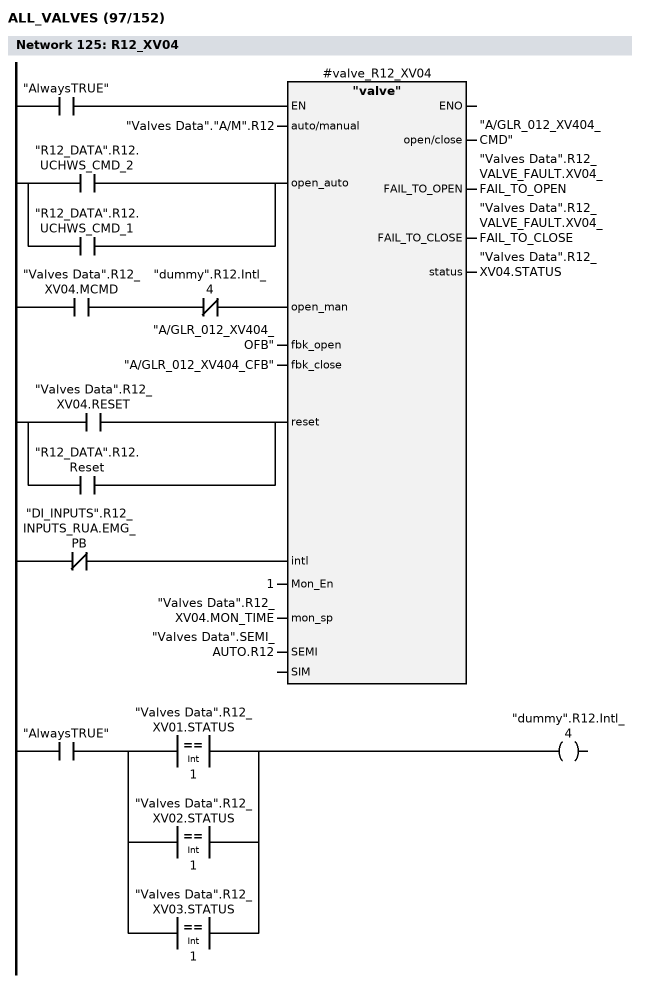
   RUNG wire#powerrail
      Contact( "AlwaysTRUE" )
      #valve_R12_XV04(open_auto := wire#w1, open_man := wire#w2, reset := wire#w3, intl := wire#w4, "auto/manual" := "Valves Data"."A/M".R12, fbk_open := "A/GLR_012_XV404_OFB", fbk_close := "A/GLR_012_XV404_CFB", Mon_En := 1, mon_sp := "Valves Data".R12_XV04.MON_TIME, SEMI := "Valves Data".SEMI_AUTO.R12, SIM :=, "open/close" => "A/GLR_012_XV404_CMD", FAIL_TO_OPEN => "Valves Data".R12_VALVE_FAULT.XV04_FAIL_TO_OPEN, FAIL_TO_CLOSE => "Valves Data".R12_VALVE_FAULT.XV04_FAIL_TO_CLOSE, status => "Valves Data".R12_XV04.STATUS)
   END_RUNG
   RUNG wire#powerrail
      Contact( "R12_DATA".R12.UCHWS_CMD_2 )
   END_RUNG wire#w1
   RUNG wire#powerrail
      Contact( "R12_DATA".R12.UCHWS_CMD_1 )
   END_RUNG wire#w1
   RUNG wire#powerrail
      Contact( "Valves Data".R12_XV04.MCMD )
      I_Contact( "dummy".R12.Intl_4 )
   END_RUNG wire#w2
   RUNG wire#powerrail
      Contact( "Valves Data".R12_XV04.RESET )
   END_RUNG wire#w3
   RUNG wire#powerrail
      Contact( "R12_DATA".R12.Reset )
   END_RUNG wire#w3
   RUNG wire#powerrail
      I_Contact( "DI_INPUTS".R12_INPUTS_RUA.EMG_PB )
   END_RUNG wire#w4
   RUNG wire#powerrail
      Contact( "AlwaysTRUE" )
      wire#w5
      { S7_Templates := "SrcType := Int" } EQ_Contact(in1 := "Valves Data".R12_XV01.STATUS, in2 := 1)
      wire#w6
      Coil( "dummy".R12.Intl_4 )
   END_RUNG
   RUNG wire#w5
      { S7_Templates := "SrcType := Int" } EQ_Contact(in1 := "Valves Data".R12_XV02.STATUS, in2 := 1)
   END_RUNG wire#w6
   RUNG wire#w5
      { S7_Templates := "SrcType := Int" } EQ_Contact(in1 := "Valves Data".R12_XV03.STATUS, in2 := 1)
   END_RUNG wire#w6
   // the same network as SCL:
   IF "AlwaysTRUE" THEN
       #valve_R12_XV04("auto/manual" := "Valves Data"."A/M".R12,   // "valve"
                       open_auto := "R12_DATA".R12.UCHWS_CMD_2 OR "R12_DATA".R12.UCHWS_CMD_1,
                       open_man := "Valves Data".R12_XV04.MCMD AND NOT "dummy".R12.Intl_4,
                       fbk_open := "A/GLR_012_XV404_OFB",
                       fbk_close := "A/GLR_012_XV404_CFB",
                       reset := "Valves Data".R12_XV04.RESET OR "R12_DATA".R12.Reset,
                       intl := NOT "DI_INPUTS".R12_INPUTS_RUA.EMG_PB,
                       Mon_En := 1,
                       mon_sp := "Valves Data".R12_XV04.MON_TIME,
                       SEMI := "Valves Data".SEMI_AUTO.R12,
                       "open/close" => "A/GLR_012_XV404_CMD",
                       FAIL_TO_OPEN => "Valves Data".R12_VALVE_FAULT.XV04_FAIL_TO_OPEN,
                       FAIL_TO_CLOSE => "Valves Data".R12_VALVE_FAULT.XV04_FAIL_TO_CLOSE,
                       status => "Valves Data".R12_XV04.STATUS);
   END_IF;
   "dummy".R12.Intl_4 := "AlwaysTRUE" AND (("Valves Data".R12_XV01.STATUS = 1) OR ("Valves Data".R12_XV02.STATUS = 1) OR ("Valves Data".R12_XV03.STATUS = 1));
END_REGION

REGION Network 126: R12_XV05
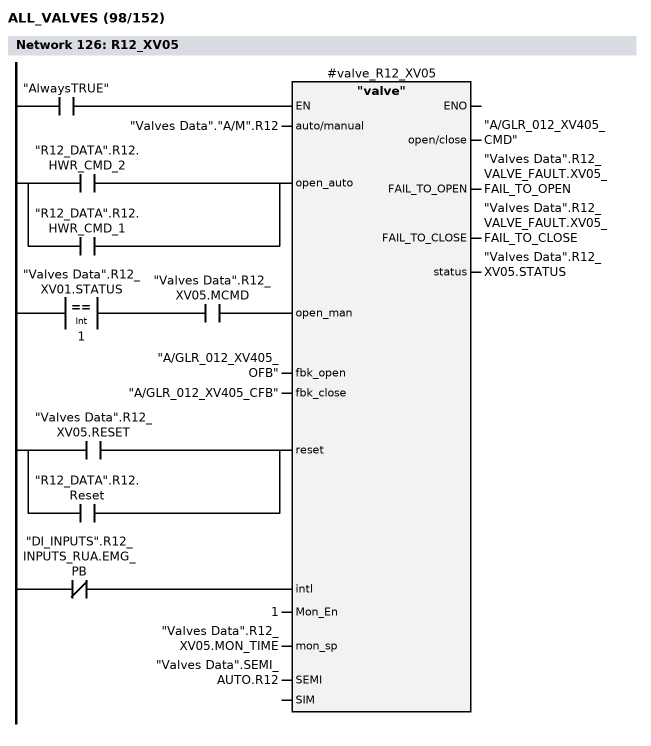
   RUNG wire#powerrail
      Contact( "AlwaysTRUE" )
      #valve_R12_XV05(open_auto := wire#w1, open_man := wire#w2, reset := wire#w3, intl := wire#w4, "auto/manual" := "Valves Data"."A/M".R12, fbk_open := "A/GLR_012_XV405_OFB", fbk_close := "A/GLR_012_XV405_CFB", Mon_En := 1, mon_sp := "Valves Data".R12_XV05.MON_TIME, SEMI := "Valves Data".SEMI_AUTO.R12, SIM :=, "open/close" => "A/GLR_012_XV405_CMD", FAIL_TO_OPEN => "Valves Data".R12_VALVE_FAULT.XV05_FAIL_TO_OPEN, FAIL_TO_CLOSE => "Valves Data".R12_VALVE_FAULT.XV05_FAIL_TO_CLOSE, status => "Valves Data".R12_XV05.STATUS)
   END_RUNG
   RUNG wire#powerrail
      Contact( "R12_DATA".R12.HWR_CMD_2 )
   END_RUNG wire#w1
   RUNG wire#powerrail
      Contact( "R12_DATA".R12.HWR_CMD_1 )
   END_RUNG wire#w1
   RUNG wire#powerrail
      { S7_Templates := "SrcType := Int" } EQ_Contact(in1 := "Valves Data".R12_XV01.STATUS, in2 := 1)
      Contact( "Valves Data".R12_XV05.MCMD )
   END_RUNG wire#w2
   RUNG wire#powerrail
      Contact( "Valves Data".R12_XV05.RESET )
   END_RUNG wire#w3
   RUNG wire#powerrail
      Contact( "R12_DATA".R12.Reset )
   END_RUNG wire#w3
   RUNG wire#powerrail
      I_Contact( "DI_INPUTS".R12_INPUTS_RUA.EMG_PB )
   END_RUNG wire#w4
   // the same network as SCL:
   IF "AlwaysTRUE" THEN
       #valve_R12_XV05("auto/manual" := "Valves Data"."A/M".R12,   // "valve"
                       open_auto := "R12_DATA".R12.HWR_CMD_2 OR "R12_DATA".R12.HWR_CMD_1,
                       open_man := ("Valves Data".R12_XV01.STATUS = 1) AND "Valves Data".R12_XV05.MCMD,
                       fbk_open := "A/GLR_012_XV405_OFB",
                       fbk_close := "A/GLR_012_XV405_CFB",
                       reset := "Valves Data".R12_XV05.RESET OR "R12_DATA".R12.Reset,
                       intl := NOT "DI_INPUTS".R12_INPUTS_RUA.EMG_PB,
                       Mon_En := 1,
                       mon_sp := "Valves Data".R12_XV05.MON_TIME,
                       SEMI := "Valves Data".SEMI_AUTO.R12,
                       "open/close" => "A/GLR_012_XV405_CMD",
                       FAIL_TO_OPEN => "Valves Data".R12_VALVE_FAULT.XV05_FAIL_TO_OPEN,
                       FAIL_TO_CLOSE => "Valves Data".R12_VALVE_FAULT.XV05_FAIL_TO_CLOSE,
                       status => "Valves Data".R12_XV05.STATUS);
   END_IF;
END_REGION

REGION Network 127: R12_XV06
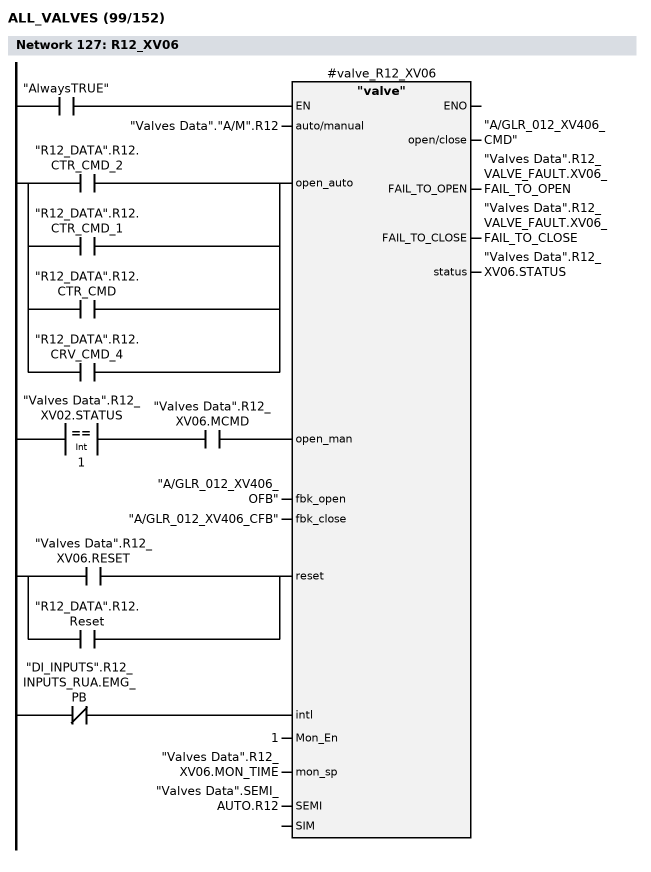
   RUNG wire#powerrail
      Contact( "AlwaysTRUE" )
      #valve_R12_XV06(open_auto := wire#w1, open_man := wire#w2, reset := wire#w3, intl := wire#w4, "auto/manual" := "Valves Data"."A/M".R12, fbk_open := "A/GLR_012_XV406_OFB", fbk_close := "A/GLR_012_XV406_CFB", Mon_En := 1, mon_sp := "Valves Data".R12_XV06.MON_TIME, SEMI := "Valves Data".SEMI_AUTO.R12, SIM :=, "open/close" => "A/GLR_012_XV406_CMD", FAIL_TO_OPEN => "Valves Data".R12_VALVE_FAULT.XV06_FAIL_TO_OPEN, FAIL_TO_CLOSE => "Valves Data".R12_VALVE_FAULT.XV06_FAIL_TO_CLOSE, status => "Valves Data".R12_XV06.STATUS)
   END_RUNG
   RUNG wire#powerrail
      Contact( "R12_DATA".R12.CTR_CMD_2 )
   END_RUNG wire#w1
   RUNG wire#powerrail
      Contact( "R12_DATA".R12.CTR_CMD_1 )
   END_RUNG wire#w1
   RUNG wire#powerrail
      Contact( "R12_DATA".R12.CTR_CMD )
   END_RUNG wire#w1
   RUNG wire#powerrail
      Contact( "R12_DATA".R12.CRV_CMD_4 )
   END_RUNG wire#w1
   RUNG wire#powerrail
      { S7_Templates := "SrcType := Int" } EQ_Contact(in1 := "Valves Data".R12_XV02.STATUS, in2 := 1)
      Contact( "Valves Data".R12_XV06.MCMD )
   END_RUNG wire#w2
   RUNG wire#powerrail
      Contact( "Valves Data".R12_XV06.RESET )
   END_RUNG wire#w3
   RUNG wire#powerrail
      Contact( "R12_DATA".R12.Reset )
   END_RUNG wire#w3
   RUNG wire#powerrail
      I_Contact( "DI_INPUTS".R12_INPUTS_RUA.EMG_PB )
   END_RUNG wire#w4
   // the same network as SCL:
   IF "AlwaysTRUE" THEN
       #valve_R12_XV06("auto/manual" := "Valves Data"."A/M".R12,   // "valve"
                       open_auto := "R12_DATA".R12.CTR_CMD_2 OR "R12_DATA".R12.CTR_CMD_1 OR "R12_DATA".R12.CTR_CMD OR "R12_DATA".R12.CRV_CMD_4,
                       open_man := ("Valves Data".R12_XV02.STATUS = 1) AND "Valves Data".R12_XV06.MCMD,
                       fbk_open := "A/GLR_012_XV406_OFB",
                       fbk_close := "A/GLR_012_XV406_CFB",
                       reset := "Valves Data".R12_XV06.RESET OR "R12_DATA".R12.Reset,
                       intl := NOT "DI_INPUTS".R12_INPUTS_RUA.EMG_PB,
                       Mon_En := 1,
                       mon_sp := "Valves Data".R12_XV06.MON_TIME,
                       SEMI := "Valves Data".SEMI_AUTO.R12,
                       "open/close" => "A/GLR_012_XV406_CMD",
                       FAIL_TO_OPEN => "Valves Data".R12_VALVE_FAULT.XV06_FAIL_TO_OPEN,
                       FAIL_TO_CLOSE => "Valves Data".R12_VALVE_FAULT.XV06_FAIL_TO_CLOSE,
                       status => "Valves Data".R12_XV06.STATUS);
   END_IF;
END_REGION

REGION Network 128: R12_XV07
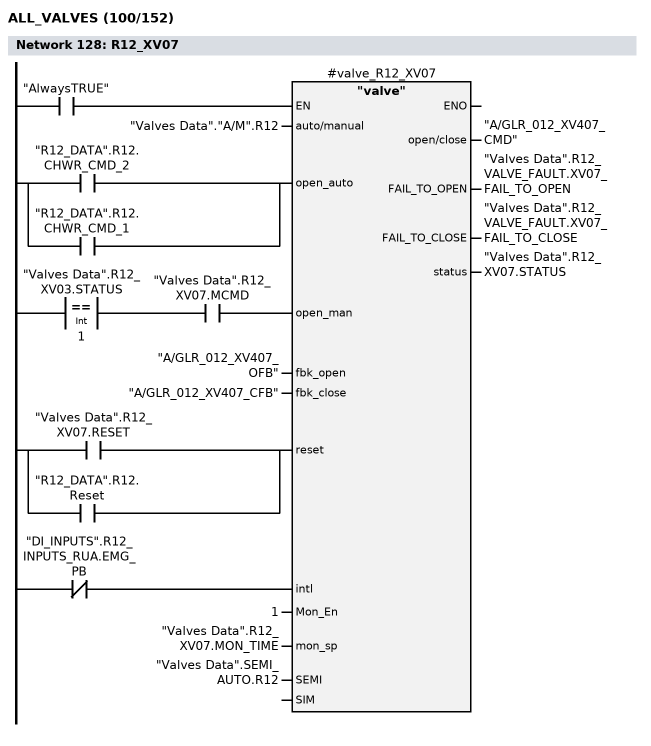
   RUNG wire#powerrail
      Contact( "AlwaysTRUE" )
      #valve_R12_XV07(open_auto := wire#w1, open_man := wire#w2, reset := wire#w3, intl := wire#w4, "auto/manual" := "Valves Data"."A/M".R12, fbk_open := "A/GLR_012_XV407_OFB", fbk_close := "A/GLR_012_XV407_CFB", Mon_En := 1, mon_sp := "Valves Data".R12_XV07.MON_TIME, SEMI := "Valves Data".SEMI_AUTO.R12, SIM :=, "open/close" => "A/GLR_012_XV407_CMD", FAIL_TO_OPEN => "Valves Data".R12_VALVE_FAULT.XV07_FAIL_TO_OPEN, FAIL_TO_CLOSE => "Valves Data".R12_VALVE_FAULT.XV07_FAIL_TO_CLOSE, status => "Valves Data".R12_XV07.STATUS)
   END_RUNG
   RUNG wire#powerrail
      Contact( "R12_DATA".R12.CHWR_CMD_2 )
   END_RUNG wire#w1
   RUNG wire#powerrail
      Contact( "R12_DATA".R12.CHWR_CMD_1 )
   END_RUNG wire#w1
   RUNG wire#powerrail
      { S7_Templates := "SrcType := Int" } EQ_Contact(in1 := "Valves Data".R12_XV03.STATUS, in2 := 1)
      Contact( "Valves Data".R12_XV07.MCMD )
   END_RUNG wire#w2
   RUNG wire#powerrail
      Contact( "Valves Data".R12_XV07.RESET )
   END_RUNG wire#w3
   RUNG wire#powerrail
      Contact( "R12_DATA".R12.Reset )
   END_RUNG wire#w3
   RUNG wire#powerrail
      I_Contact( "DI_INPUTS".R12_INPUTS_RUA.EMG_PB )
   END_RUNG wire#w4
   // the same network as SCL:
   IF "AlwaysTRUE" THEN
       #valve_R12_XV07("auto/manual" := "Valves Data"."A/M".R12,   // "valve"
                       open_auto := "R12_DATA".R12.CHWR_CMD_2 OR "R12_DATA".R12.CHWR_CMD_1,
                       open_man := ("Valves Data".R12_XV03.STATUS = 1) AND "Valves Data".R12_XV07.MCMD,
                       fbk_open := "A/GLR_012_XV407_OFB",
                       fbk_close := "A/GLR_012_XV407_CFB",
                       reset := "Valves Data".R12_XV07.RESET OR "R12_DATA".R12.Reset,
                       intl := NOT "DI_INPUTS".R12_INPUTS_RUA.EMG_PB,
                       Mon_En := 1,
                       mon_sp := "Valves Data".R12_XV07.MON_TIME,
                       SEMI := "Valves Data".SEMI_AUTO.R12,
                       "open/close" => "A/GLR_012_XV407_CMD",
                       FAIL_TO_OPEN => "Valves Data".R12_VALVE_FAULT.XV07_FAIL_TO_OPEN,
                       FAIL_TO_CLOSE => "Valves Data".R12_VALVE_FAULT.XV07_FAIL_TO_CLOSE,
                       status => "Valves Data".R12_XV07.STATUS);
   END_IF;
END_REGION

REGION Network 129: R12_XV08
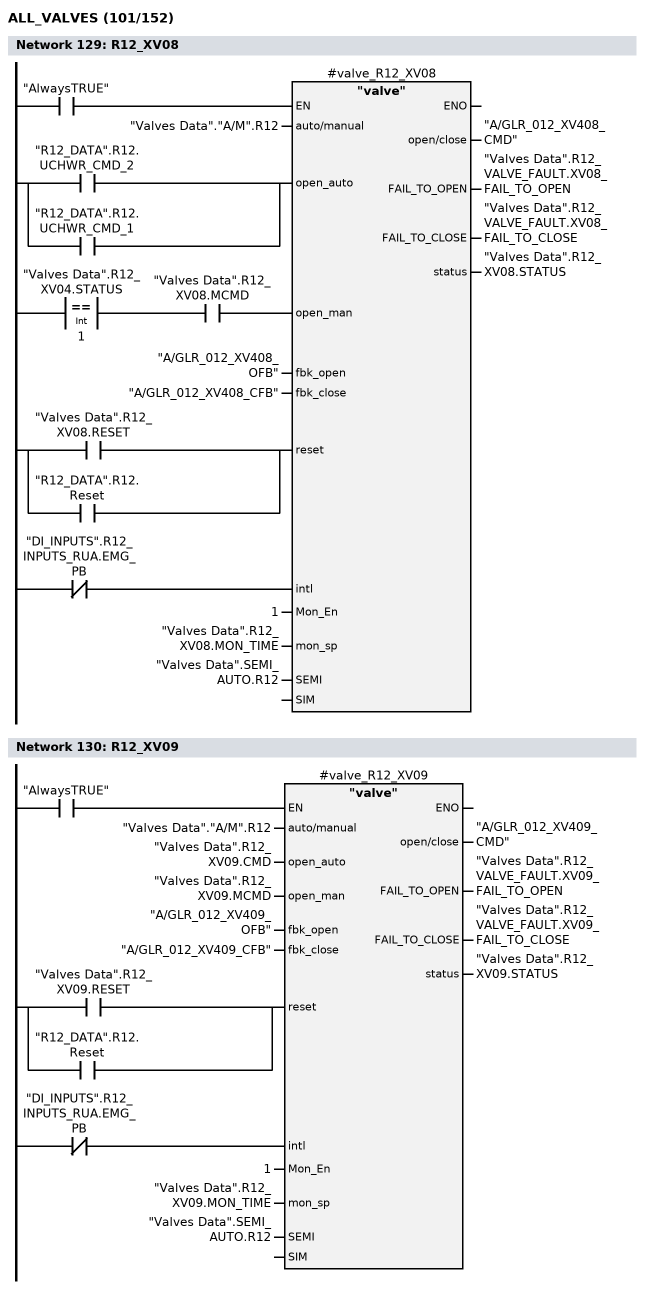
   RUNG wire#powerrail
      Contact( "AlwaysTRUE" )
      #valve_R12_XV08(open_auto := wire#w1, open_man := wire#w2, reset := wire#w3, intl := wire#w4, "auto/manual" := "Valves Data"."A/M".R12, fbk_open := "A/GLR_012_XV408_OFB", fbk_close := "A/GLR_012_XV408_CFB", Mon_En := 1, mon_sp := "Valves Data".R12_XV08.MON_TIME, SEMI := "Valves Data".SEMI_AUTO.R12, SIM :=, "open/close" => "A/GLR_012_XV408_CMD", FAIL_TO_OPEN => "Valves Data".R12_VALVE_FAULT.XV08_FAIL_TO_OPEN, FAIL_TO_CLOSE => "Valves Data".R12_VALVE_FAULT.XV08_FAIL_TO_CLOSE, status => "Valves Data".R12_XV08.STATUS)
   END_RUNG
   RUNG wire#powerrail
      Contact( "R12_DATA".R12.UCHWR_CMD_2 )
   END_RUNG wire#w1
   RUNG wire#powerrail
      Contact( "R12_DATA".R12.UCHWR_CMD_1 )
   END_RUNG wire#w1
   RUNG wire#powerrail
      { S7_Templates := "SrcType := Int" } EQ_Contact(in1 := "Valves Data".R12_XV04.STATUS, in2 := 1)
      Contact( "Valves Data".R12_XV08.MCMD )
   END_RUNG wire#w2
   RUNG wire#powerrail
      Contact( "Valves Data".R12_XV08.RESET )
   END_RUNG wire#w3
   RUNG wire#powerrail
      Contact( "R12_DATA".R12.Reset )
   END_RUNG wire#w3
   RUNG wire#powerrail
      I_Contact( "DI_INPUTS".R12_INPUTS_RUA.EMG_PB )
   END_RUNG wire#w4
   // the same network as SCL:
   IF "AlwaysTRUE" THEN
       #valve_R12_XV08("auto/manual" := "Valves Data"."A/M".R12,   // "valve"
                       open_auto := "R12_DATA".R12.UCHWR_CMD_2 OR "R12_DATA".R12.UCHWR_CMD_1,
                       open_man := ("Valves Data".R12_XV04.STATUS = 1) AND "Valves Data".R12_XV08.MCMD,
                       fbk_open := "A/GLR_012_XV408_OFB",
                       fbk_close := "A/GLR_012_XV408_CFB",
                       reset := "Valves Data".R12_XV08.RESET OR "R12_DATA".R12.Reset,
                       intl := NOT "DI_INPUTS".R12_INPUTS_RUA.EMG_PB,
                       Mon_En := 1,
                       mon_sp := "Valves Data".R12_XV08.MON_TIME,
                       SEMI := "Valves Data".SEMI_AUTO.R12,
                       "open/close" => "A/GLR_012_XV408_CMD",
                       FAIL_TO_OPEN => "Valves Data".R12_VALVE_FAULT.XV08_FAIL_TO_OPEN,
                       FAIL_TO_CLOSE => "Valves Data".R12_VALVE_FAULT.XV08_FAIL_TO_CLOSE,
                       status => "Valves Data".R12_XV08.STATUS);
   END_IF;
END_REGION

REGION Network 130: R12_XV09
   RUNG wire#powerrail
      Contact( "AlwaysTRUE" )
      #valve_R12_XV09(reset := wire#w1, intl := wire#w2, "auto/manual" := "Valves Data"."A/M".R12, open_auto := "Valves Data".R12_XV09.CMD, open_man := "Valves Data".R12_XV09.MCMD, fbk_open := "A/GLR_012_XV409_OFB", fbk_close := "A/GLR_012_XV409_CFB", Mon_En := 1, mon_sp := "Valves Data".R12_XV09.MON_TIME, SEMI := "Valves Data".SEMI_AUTO.R12, SIM :=, "open/close" => "A/GLR_012_XV409_CMD", FAIL_TO_OPEN => "Valves Data".R12_VALVE_FAULT.XV09_FAIL_TO_OPEN, FAIL_TO_CLOSE => "Valves Data".R12_VALVE_FAULT.XV09_FAIL_TO_CLOSE, status => "Valves Data".R12_XV09.STATUS)
   END_RUNG
   RUNG wire#powerrail
      Contact( "Valves Data".R12_XV09.RESET )
   END_RUNG wire#w1
   RUNG wire#powerrail
      Contact( "R12_DATA".R12.Reset )
   END_RUNG wire#w1
   RUNG wire#powerrail
      I_Contact( "DI_INPUTS".R12_INPUTS_RUA.EMG_PB )
   END_RUNG wire#w2
   // the same network as SCL:
   IF "AlwaysTRUE" THEN
       #valve_R12_XV09("auto/manual" := "Valves Data"."A/M".R12,   // "valve"
                       open_auto := "Valves Data".R12_XV09.CMD,
                       open_man := "Valves Data".R12_XV09.MCMD,
                       fbk_open := "A/GLR_012_XV409_OFB",
                       fbk_close := "A/GLR_012_XV409_CFB",
                       reset := "Valves Data".R12_XV09.RESET OR "R12_DATA".R12.Reset,
                       intl := NOT "DI_INPUTS".R12_INPUTS_RUA.EMG_PB,
                       Mon_En := 1,
                       mon_sp := "Valves Data".R12_XV09.MON_TIME,
                       SEMI := "Valves Data".SEMI_AUTO.R12,
                       "open/close" => "A/GLR_012_XV409_CMD",
                       FAIL_TO_OPEN => "Valves Data".R12_VALVE_FAULT.XV09_FAIL_TO_OPEN,
                       FAIL_TO_CLOSE => "Valves Data".R12_VALVE_FAULT.XV09_FAIL_TO_CLOSE,
                       status => "Valves Data".R12_XV09.STATUS);
   END_IF;
END_REGION

REGION Network 131: ****REACTOR_13****
END_REGION

REGION Network 132: R13_XV01
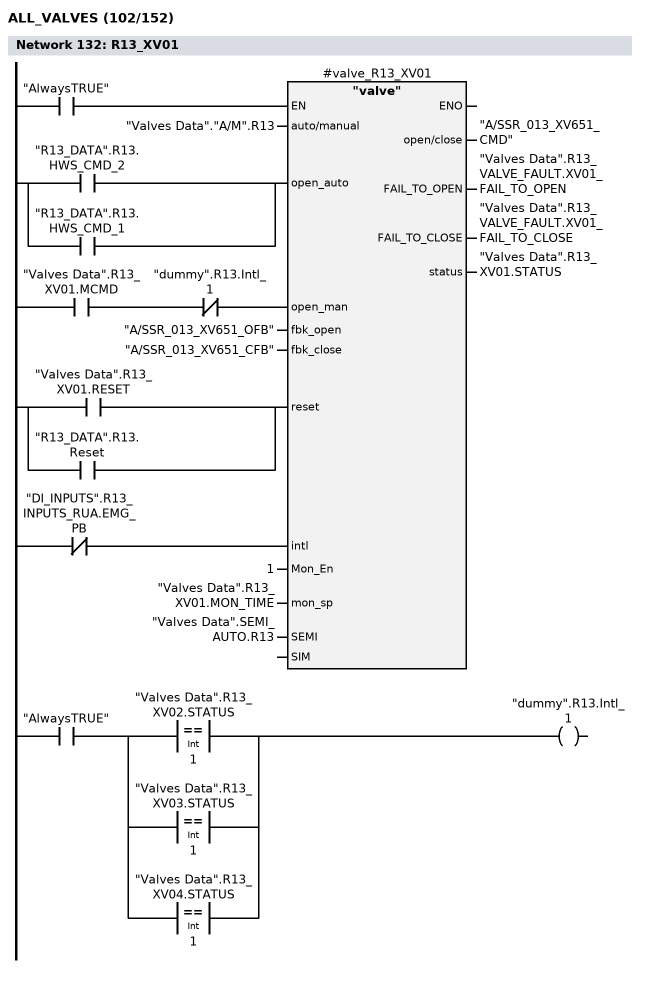
   RUNG wire#powerrail
      Contact( "AlwaysTRUE" )
      #valve_R13_XV01(open_auto := wire#w1, open_man := wire#w2, reset := wire#w3, intl := wire#w4, "auto/manual" := "Valves Data"."A/M".R13, fbk_open := "A/SSR_013_XV651_OFB", fbk_close := "A/SSR_013_XV651_CFB", Mon_En := 1, mon_sp := "Valves Data".R13_XV01.MON_TIME, SEMI := "Valves Data".SEMI_AUTO.R13, SIM :=, "open/close" => "A/SSR_013_XV651_CMD", FAIL_TO_OPEN => "Valves Data".R13_VALVE_FAULT.XV01_FAIL_TO_OPEN, FAIL_TO_CLOSE => "Valves Data".R13_VALVE_FAULT.XV01_FAIL_TO_CLOSE, status => "Valves Data".R13_XV01.STATUS)
   END_RUNG
   RUNG wire#powerrail
      Contact( "R13_DATA".R13.HWS_CMD_2 )
   END_RUNG wire#w1
   RUNG wire#powerrail
      Contact( "R13_DATA".R13.HWS_CMD_1 )
   END_RUNG wire#w1
   RUNG wire#powerrail
      Contact( "Valves Data".R13_XV01.MCMD )
      I_Contact( "dummy".R13.Intl_1 )
   END_RUNG wire#w2
   RUNG wire#powerrail
      Contact( "Valves Data".R13_XV01.RESET )
   END_RUNG wire#w3
   RUNG wire#powerrail
      Contact( "R13_DATA".R13.Reset )
   END_RUNG wire#w3
   RUNG wire#powerrail
      I_Contact( "DI_INPUTS".R13_INPUTS_RUA.EMG_PB )
   END_RUNG wire#w4
   RUNG wire#powerrail
      Contact( "AlwaysTRUE" )
      wire#w5
      { S7_Templates := "SrcType := Int" } EQ_Contact(in1 := "Valves Data".R13_XV02.STATUS, in2 := 1)
      wire#w6
      Coil( "dummy".R13.Intl_1 )
   END_RUNG
   RUNG wire#w5
      { S7_Templates := "SrcType := Int" } EQ_Contact(in1 := "Valves Data".R13_XV03.STATUS, in2 := 1)
   END_RUNG wire#w6
   RUNG wire#w5
      { S7_Templates := "SrcType := Int" } EQ_Contact(in1 := "Valves Data".R13_XV04.STATUS, in2 := 1)
   END_RUNG wire#w6
   // the same network as SCL:
   IF "AlwaysTRUE" THEN
       #valve_R13_XV01("auto/manual" := "Valves Data"."A/M".R13,   // "valve"
                       open_auto := "R13_DATA".R13.HWS_CMD_2 OR "R13_DATA".R13.HWS_CMD_1,
                       open_man := "Valves Data".R13_XV01.MCMD AND NOT "dummy".R13.Intl_1,
                       fbk_open := "A/SSR_013_XV651_OFB",
                       fbk_close := "A/SSR_013_XV651_CFB",
                       reset := "Valves Data".R13_XV01.RESET OR "R13_DATA".R13.Reset,
                       intl := NOT "DI_INPUTS".R13_INPUTS_RUA.EMG_PB,
                       Mon_En := 1,
                       mon_sp := "Valves Data".R13_XV01.MON_TIME,
                       SEMI := "Valves Data".SEMI_AUTO.R13,
                       "open/close" => "A/SSR_013_XV651_CMD",
                       FAIL_TO_OPEN => "Valves Data".R13_VALVE_FAULT.XV01_FAIL_TO_OPEN,
                       FAIL_TO_CLOSE => "Valves Data".R13_VALVE_FAULT.XV01_FAIL_TO_CLOSE,
                       status => "Valves Data".R13_XV01.STATUS);
   END_IF;
   "dummy".R13.Intl_1 := "AlwaysTRUE" AND (("Valves Data".R13_XV02.STATUS = 1) OR ("Valves Data".R13_XV03.STATUS = 1) OR ("Valves Data".R13_XV04.STATUS = 1));
END_REGION

REGION Network 133: R13_XV02
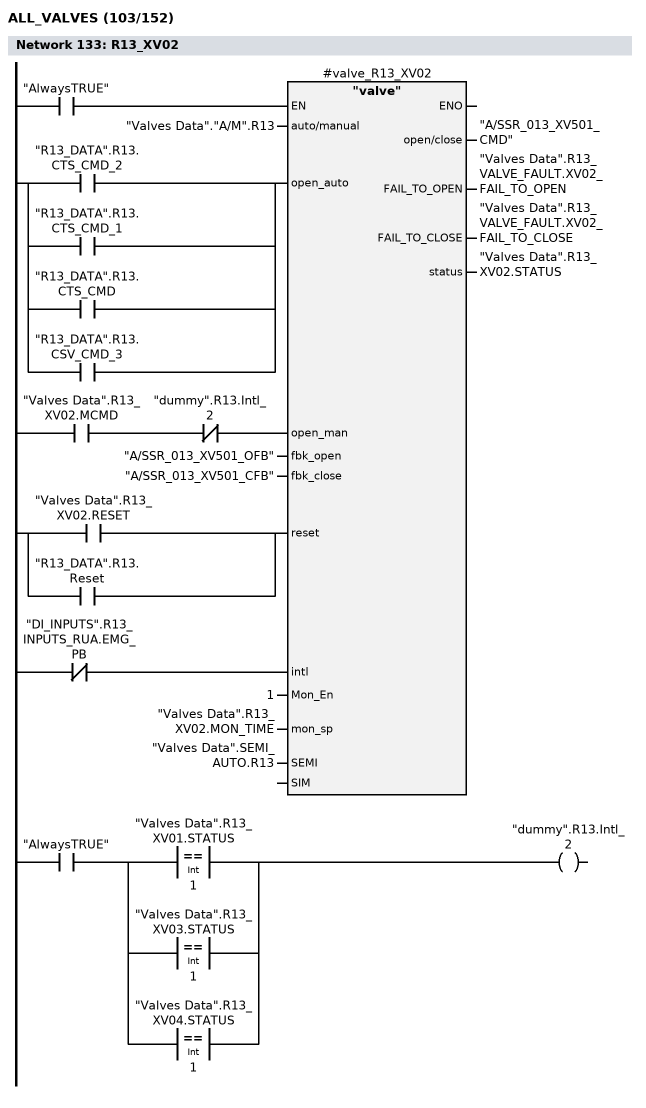
   RUNG wire#powerrail
      Contact( "AlwaysTRUE" )
      #valve_R13_XV02(open_auto := wire#w1, open_man := wire#w2, reset := wire#w3, intl := wire#w4, "auto/manual" := "Valves Data"."A/M".R13, fbk_open := "A/SSR_013_XV501_OFB", fbk_close := "A/SSR_013_XV501_CFB", Mon_En := 1, mon_sp := "Valves Data".R13_XV02.MON_TIME, SEMI := "Valves Data".SEMI_AUTO.R13, SIM :=, "open/close" => "A/SSR_013_XV501_CMD", FAIL_TO_OPEN => "Valves Data".R13_VALVE_FAULT.XV02_FAIL_TO_OPEN, FAIL_TO_CLOSE => "Valves Data".R13_VALVE_FAULT.XV02_FAIL_TO_CLOSE, status => "Valves Data".R13_XV02.STATUS)
   END_RUNG
   RUNG wire#powerrail
      Contact( "R13_DATA".R13.CTS_CMD_2 )
   END_RUNG wire#w1
   RUNG wire#powerrail
      Contact( "R13_DATA".R13.CTS_CMD_1 )
   END_RUNG wire#w1
   RUNG wire#powerrail
      Contact( "R13_DATA".R13.CTS_CMD )
   END_RUNG wire#w1
   RUNG wire#powerrail
      Contact( "R13_DATA".R13.CSV_CMD_3 )
   END_RUNG wire#w1
   RUNG wire#powerrail
      Contact( "Valves Data".R13_XV02.MCMD )
      I_Contact( "dummy".R13.Intl_2 )
   END_RUNG wire#w2
   RUNG wire#powerrail
      Contact( "Valves Data".R13_XV02.RESET )
   END_RUNG wire#w3
   RUNG wire#powerrail
      Contact( "R13_DATA".R13.Reset )
   END_RUNG wire#w3
   RUNG wire#powerrail
      I_Contact( "DI_INPUTS".R13_INPUTS_RUA.EMG_PB )
   END_RUNG wire#w4
   RUNG wire#powerrail
      Contact( "AlwaysTRUE" )
      wire#w5
      { S7_Templates := "SrcType := Int" } EQ_Contact(in1 := "Valves Data".R13_XV01.STATUS, in2 := 1)
      wire#w6
      Coil( "dummy".R13.Intl_2 )
   END_RUNG
   RUNG wire#w5
      { S7_Templates := "SrcType := Int" } EQ_Contact(in1 := "Valves Data".R13_XV03.STATUS, in2 := 1)
   END_RUNG wire#w6
   RUNG wire#w5
      { S7_Templates := "SrcType := Int" } EQ_Contact(in1 := "Valves Data".R13_XV04.STATUS, in2 := 1)
   END_RUNG wire#w6
   // the same network as SCL:
   IF "AlwaysTRUE" THEN
       #valve_R13_XV02("auto/manual" := "Valves Data"."A/M".R13,   // "valve"
                       open_auto := "R13_DATA".R13.CTS_CMD_2 OR "R13_DATA".R13.CTS_CMD_1 OR "R13_DATA".R13.CTS_CMD OR "R13_DATA".R13.CSV_CMD_3,
                       open_man := "Valves Data".R13_XV02.MCMD AND NOT "dummy".R13.Intl_2,
                       fbk_open := "A/SSR_013_XV501_OFB",
                       fbk_close := "A/SSR_013_XV501_CFB",
                       reset := "Valves Data".R13_XV02.RESET OR "R13_DATA".R13.Reset,
                       intl := NOT "DI_INPUTS".R13_INPUTS_RUA.EMG_PB,
                       Mon_En := 1,
                       mon_sp := "Valves Data".R13_XV02.MON_TIME,
                       SEMI := "Valves Data".SEMI_AUTO.R13,
                       "open/close" => "A/SSR_013_XV501_CMD",
                       FAIL_TO_OPEN => "Valves Data".R13_VALVE_FAULT.XV02_FAIL_TO_OPEN,
                       FAIL_TO_CLOSE => "Valves Data".R13_VALVE_FAULT.XV02_FAIL_TO_CLOSE,
                       status => "Valves Data".R13_XV02.STATUS);
   END_IF;
   "dummy".R13.Intl_2 := "AlwaysTRUE" AND (("Valves Data".R13_XV01.STATUS = 1) OR ("Valves Data".R13_XV03.STATUS = 1) OR ("Valves Data".R13_XV04.STATUS = 1));
END_REGION

REGION Network 134: R13_XV03
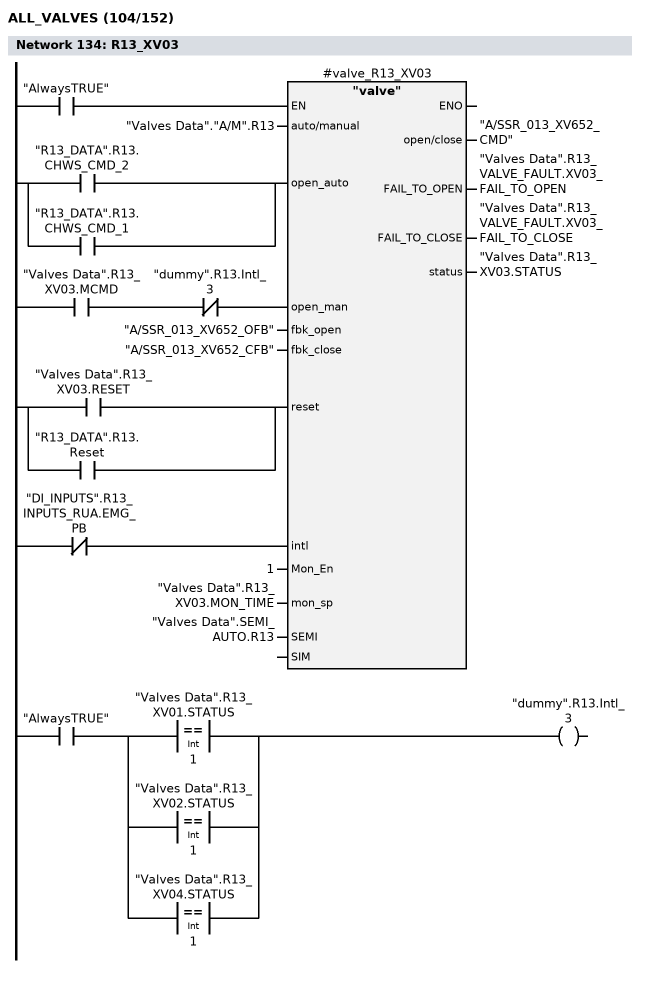
   RUNG wire#powerrail
      Contact( "AlwaysTRUE" )
      #valve_R13_XV03(open_auto := wire#w1, open_man := wire#w2, reset := wire#w3, intl := wire#w4, "auto/manual" := "Valves Data"."A/M".R13, fbk_open := "A/SSR_013_XV652_OFB", fbk_close := "A/SSR_013_XV652_CFB", Mon_En := 1, mon_sp := "Valves Data".R13_XV03.MON_TIME, SEMI := "Valves Data".SEMI_AUTO.R13, SIM :=, "open/close" => "A/SSR_013_XV652_CMD", FAIL_TO_OPEN => "Valves Data".R13_VALVE_FAULT.XV03_FAIL_TO_OPEN, FAIL_TO_CLOSE => "Valves Data".R13_VALVE_FAULT.XV03_FAIL_TO_CLOSE, status => "Valves Data".R13_XV03.STATUS)
   END_RUNG
   RUNG wire#powerrail
      Contact( "R13_DATA".R13.CHWS_CMD_2 )
   END_RUNG wire#w1
   RUNG wire#powerrail
      Contact( "R13_DATA".R13.CHWS_CMD_1 )
   END_RUNG wire#w1
   RUNG wire#powerrail
      Contact( "Valves Data".R13_XV03.MCMD )
      I_Contact( "dummy".R13.Intl_3 )
   END_RUNG wire#w2
   RUNG wire#powerrail
      Contact( "Valves Data".R13_XV03.RESET )
   END_RUNG wire#w3
   RUNG wire#powerrail
      Contact( "R13_DATA".R13.Reset )
   END_RUNG wire#w3
   RUNG wire#powerrail
      I_Contact( "DI_INPUTS".R13_INPUTS_RUA.EMG_PB )
   END_RUNG wire#w4
   RUNG wire#powerrail
      Contact( "AlwaysTRUE" )
      wire#w5
      { S7_Templates := "SrcType := Int" } EQ_Contact(in1 := "Valves Data".R13_XV01.STATUS, in2 := 1)
      wire#w6
      Coil( "dummy".R13.Intl_3 )
   END_RUNG
   RUNG wire#w5
      { S7_Templates := "SrcType := Int" } EQ_Contact(in1 := "Valves Data".R13_XV02.STATUS, in2 := 1)
   END_RUNG wire#w6
   RUNG wire#w5
      { S7_Templates := "SrcType := Int" } EQ_Contact(in1 := "Valves Data".R13_XV04.STATUS, in2 := 1)
   END_RUNG wire#w6
   // the same network as SCL:
   IF "AlwaysTRUE" THEN
       #valve_R13_XV03("auto/manual" := "Valves Data"."A/M".R13,   // "valve"
                       open_auto := "R13_DATA".R13.CHWS_CMD_2 OR "R13_DATA".R13.CHWS_CMD_1,
                       open_man := "Valves Data".R13_XV03.MCMD AND NOT "dummy".R13.Intl_3,
                       fbk_open := "A/SSR_013_XV652_OFB",
                       fbk_close := "A/SSR_013_XV652_CFB",
                       reset := "Valves Data".R13_XV03.RESET OR "R13_DATA".R13.Reset,
                       intl := NOT "DI_INPUTS".R13_INPUTS_RUA.EMG_PB,
                       Mon_En := 1,
                       mon_sp := "Valves Data".R13_XV03.MON_TIME,
                       SEMI := "Valves Data".SEMI_AUTO.R13,
                       "open/close" => "A/SSR_013_XV652_CMD",
                       FAIL_TO_OPEN => "Valves Data".R13_VALVE_FAULT.XV03_FAIL_TO_OPEN,
                       FAIL_TO_CLOSE => "Valves Data".R13_VALVE_FAULT.XV03_FAIL_TO_CLOSE,
                       status => "Valves Data".R13_XV03.STATUS);
   END_IF;
   "dummy".R13.Intl_3 := "AlwaysTRUE" AND (("Valves Data".R13_XV01.STATUS = 1) OR ("Valves Data".R13_XV02.STATUS = 1) OR ("Valves Data".R13_XV04.STATUS = 1));
END_REGION

REGION Network 135: R13_XV04
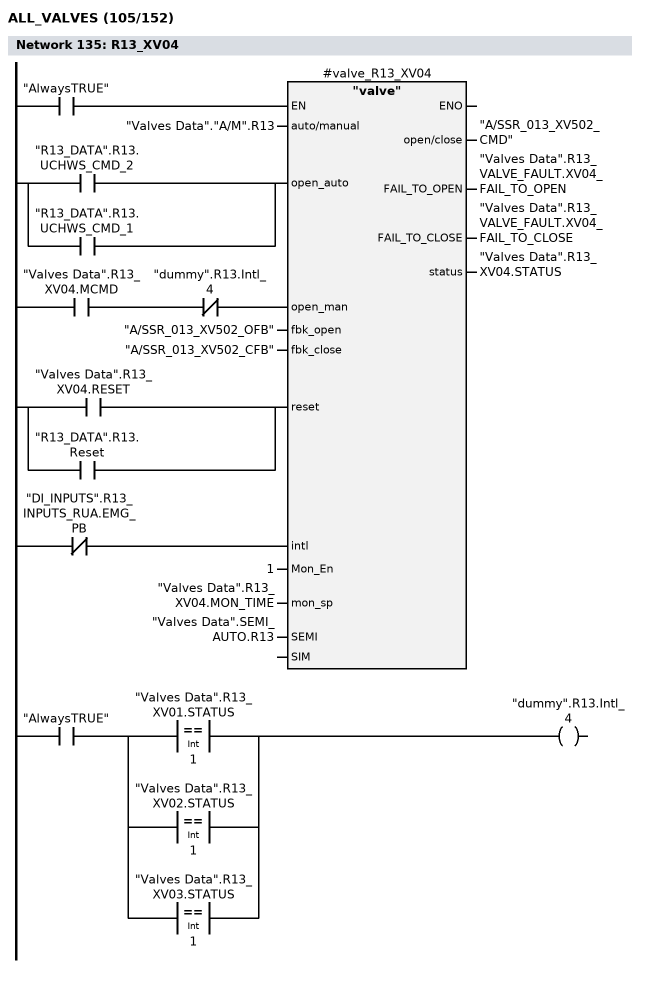
   RUNG wire#powerrail
      Contact( "AlwaysTRUE" )
      #valve_R13_XV04(open_auto := wire#w1, open_man := wire#w2, reset := wire#w3, intl := wire#w4, "auto/manual" := "Valves Data"."A/M".R13, fbk_open := "A/SSR_013_XV502_OFB", fbk_close := "A/SSR_013_XV502_CFB", Mon_En := 1, mon_sp := "Valves Data".R13_XV04.MON_TIME, SEMI := "Valves Data".SEMI_AUTO.R13, SIM :=, "open/close" => "A/SSR_013_XV502_CMD", FAIL_TO_OPEN => "Valves Data".R13_VALVE_FAULT.XV04_FAIL_TO_OPEN, FAIL_TO_CLOSE => "Valves Data".R13_VALVE_FAULT.XV04_FAIL_TO_CLOSE, status => "Valves Data".R13_XV04.STATUS)
   END_RUNG
   RUNG wire#powerrail
      Contact( "R13_DATA".R13.UCHWS_CMD_2 )
   END_RUNG wire#w1
   RUNG wire#powerrail
      Contact( "R13_DATA".R13.UCHWS_CMD_1 )
   END_RUNG wire#w1
   RUNG wire#powerrail
      Contact( "Valves Data".R13_XV04.MCMD )
      I_Contact( "dummy".R13.Intl_4 )
   END_RUNG wire#w2
   RUNG wire#powerrail
      Contact( "Valves Data".R13_XV04.RESET )
   END_RUNG wire#w3
   RUNG wire#powerrail
      Contact( "R13_DATA".R13.Reset )
   END_RUNG wire#w3
   RUNG wire#powerrail
      I_Contact( "DI_INPUTS".R13_INPUTS_RUA.EMG_PB )
   END_RUNG wire#w4
   RUNG wire#powerrail
      Contact( "AlwaysTRUE" )
      wire#w5
      { S7_Templates := "SrcType := Int" } EQ_Contact(in1 := "Valves Data".R13_XV01.STATUS, in2 := 1)
      wire#w6
      Coil( "dummy".R13.Intl_4 )
   END_RUNG
   RUNG wire#w5
      { S7_Templates := "SrcType := Int" } EQ_Contact(in1 := "Valves Data".R13_XV02.STATUS, in2 := 1)
   END_RUNG wire#w6
   RUNG wire#w5
      { S7_Templates := "SrcType := Int" } EQ_Contact(in1 := "Valves Data".R13_XV03.STATUS, in2 := 1)
   END_RUNG wire#w6
   // the same network as SCL:
   IF "AlwaysTRUE" THEN
       #valve_R13_XV04("auto/manual" := "Valves Data"."A/M".R13,   // "valve"
                       open_auto := "R13_DATA".R13.UCHWS_CMD_2 OR "R13_DATA".R13.UCHWS_CMD_1,
                       open_man := "Valves Data".R13_XV04.MCMD AND NOT "dummy".R13.Intl_4,
                       fbk_open := "A/SSR_013_XV502_OFB",
                       fbk_close := "A/SSR_013_XV502_CFB",
                       reset := "Valves Data".R13_XV04.RESET OR "R13_DATA".R13.Reset,
                       intl := NOT "DI_INPUTS".R13_INPUTS_RUA.EMG_PB,
                       Mon_En := 1,
                       mon_sp := "Valves Data".R13_XV04.MON_TIME,
                       SEMI := "Valves Data".SEMI_AUTO.R13,
                       "open/close" => "A/SSR_013_XV502_CMD",
                       FAIL_TO_OPEN => "Valves Data".R13_VALVE_FAULT.XV04_FAIL_TO_OPEN,
                       FAIL_TO_CLOSE => "Valves Data".R13_VALVE_FAULT.XV04_FAIL_TO_CLOSE,
                       status => "Valves Data".R13_XV04.STATUS);
   END_IF;
   "dummy".R13.Intl_4 := "AlwaysTRUE" AND (("Valves Data".R13_XV01.STATUS = 1) OR ("Valves Data".R13_XV02.STATUS = 1) OR ("Valves Data".R13_XV03.STATUS = 1));
END_REGION

REGION Network 136: R13_XV05
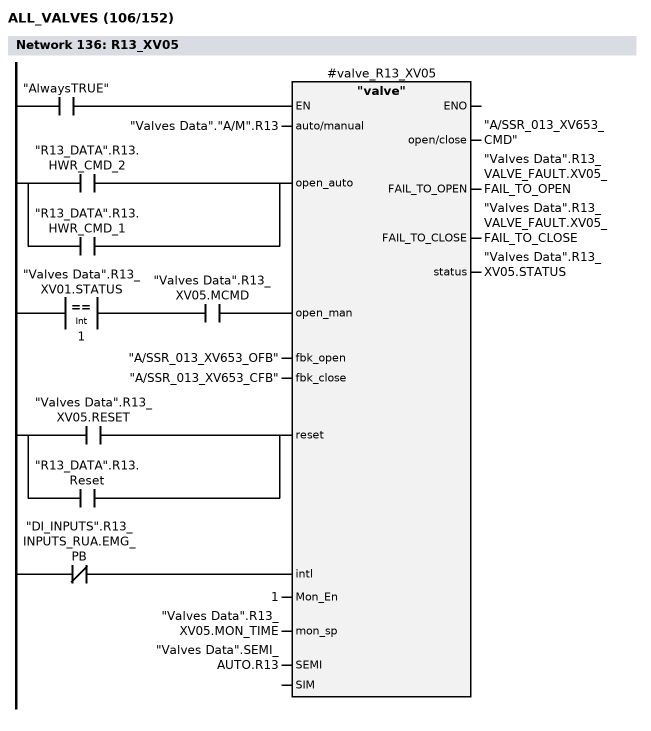
   RUNG wire#powerrail
      Contact( "AlwaysTRUE" )
      #valve_R13_XV05(open_auto := wire#w1, open_man := wire#w2, reset := wire#w3, intl := wire#w4, "auto/manual" := "Valves Data"."A/M".R13, fbk_open := "A/SSR_013_XV653_OFB", fbk_close := "A/SSR_013_XV653_CFB", Mon_En := 1, mon_sp := "Valves Data".R13_XV05.MON_TIME, SEMI := "Valves Data".SEMI_AUTO.R13, SIM :=, "open/close" => "A/SSR_013_XV653_CMD", FAIL_TO_OPEN => "Valves Data".R13_VALVE_FAULT.XV05_FAIL_TO_OPEN, FAIL_TO_CLOSE => "Valves Data".R13_VALVE_FAULT.XV05_FAIL_TO_CLOSE, status => "Valves Data".R13_XV05.STATUS)
   END_RUNG
   RUNG wire#powerrail
      Contact( "R13_DATA".R13.HWR_CMD_2 )
   END_RUNG wire#w1
   RUNG wire#powerrail
      Contact( "R13_DATA".R13.HWR_CMD_1 )
   END_RUNG wire#w1
   RUNG wire#powerrail
      { S7_Templates := "SrcType := Int" } EQ_Contact(in1 := "Valves Data".R13_XV01.STATUS, in2 := 1)
      Contact( "Valves Data".R13_XV05.MCMD )
   END_RUNG wire#w2
   RUNG wire#powerrail
      Contact( "Valves Data".R13_XV05.RESET )
   END_RUNG wire#w3
   RUNG wire#powerrail
      Contact( "R13_DATA".R13.Reset )
   END_RUNG wire#w3
   RUNG wire#powerrail
      I_Contact( "DI_INPUTS".R13_INPUTS_RUA.EMG_PB )
   END_RUNG wire#w4
   // the same network as SCL:
   IF "AlwaysTRUE" THEN
       #valve_R13_XV05("auto/manual" := "Valves Data"."A/M".R13,   // "valve"
                       open_auto := "R13_DATA".R13.HWR_CMD_2 OR "R13_DATA".R13.HWR_CMD_1,
                       open_man := ("Valves Data".R13_XV01.STATUS = 1) AND "Valves Data".R13_XV05.MCMD,
                       fbk_open := "A/SSR_013_XV653_OFB",
                       fbk_close := "A/SSR_013_XV653_CFB",
                       reset := "Valves Data".R13_XV05.RESET OR "R13_DATA".R13.Reset,
                       intl := NOT "DI_INPUTS".R13_INPUTS_RUA.EMG_PB,
                       Mon_En := 1,
                       mon_sp := "Valves Data".R13_XV05.MON_TIME,
                       SEMI := "Valves Data".SEMI_AUTO.R13,
                       "open/close" => "A/SSR_013_XV653_CMD",
                       FAIL_TO_OPEN => "Valves Data".R13_VALVE_FAULT.XV05_FAIL_TO_OPEN,
                       FAIL_TO_CLOSE => "Valves Data".R13_VALVE_FAULT.XV05_FAIL_TO_CLOSE,
                       status => "Valves Data".R13_XV05.STATUS);
   END_IF;
END_REGION

REGION Network 137: R13_XV06
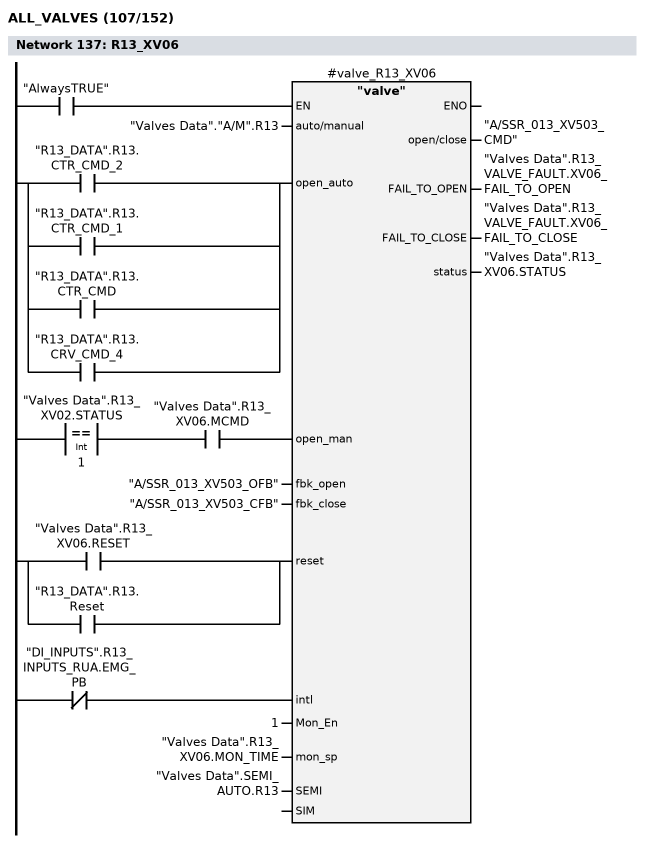
   RUNG wire#powerrail
      Contact( "AlwaysTRUE" )
      #valve_R13_XV06(open_auto := wire#w1, open_man := wire#w2, reset := wire#w3, intl := wire#w4, "auto/manual" := "Valves Data"."A/M".R13, fbk_open := "A/SSR_013_XV503_OFB", fbk_close := "A/SSR_013_XV503_CFB", Mon_En := 1, mon_sp := "Valves Data".R13_XV06.MON_TIME, SEMI := "Valves Data".SEMI_AUTO.R13, SIM :=, "open/close" => "A/SSR_013_XV503_CMD", FAIL_TO_OPEN => "Valves Data".R13_VALVE_FAULT.XV06_FAIL_TO_OPEN, FAIL_TO_CLOSE => "Valves Data".R13_VALVE_FAULT.XV06_FAIL_TO_CLOSE, status => "Valves Data".R13_XV06.STATUS)
   END_RUNG
   RUNG wire#powerrail
      Contact( "R13_DATA".R13.CTR_CMD_2 )
   END_RUNG wire#w1
   RUNG wire#powerrail
      Contact( "R13_DATA".R13.CTR_CMD_1 )
   END_RUNG wire#w1
   RUNG wire#powerrail
      Contact( "R13_DATA".R13.CTR_CMD )
   END_RUNG wire#w1
   RUNG wire#powerrail
      Contact( "R13_DATA".R13.CRV_CMD_4 )
   END_RUNG wire#w1
   RUNG wire#powerrail
      { S7_Templates := "SrcType := Int" } EQ_Contact(in1 := "Valves Data".R13_XV02.STATUS, in2 := 1)
      Contact( "Valves Data".R13_XV06.MCMD )
   END_RUNG wire#w2
   RUNG wire#powerrail
      Contact( "Valves Data".R13_XV06.RESET )
   END_RUNG wire#w3
   RUNG wire#powerrail
      Contact( "R13_DATA".R13.Reset )
   END_RUNG wire#w3
   RUNG wire#powerrail
      I_Contact( "DI_INPUTS".R13_INPUTS_RUA.EMG_PB )
   END_RUNG wire#w4
   // the same network as SCL:
   IF "AlwaysTRUE" THEN
       #valve_R13_XV06("auto/manual" := "Valves Data"."A/M".R13,   // "valve"
                       open_auto := "R13_DATA".R13.CTR_CMD_2 OR "R13_DATA".R13.CTR_CMD_1 OR "R13_DATA".R13.CTR_CMD OR "R13_DATA".R13.CRV_CMD_4,
                       open_man := ("Valves Data".R13_XV02.STATUS = 1) AND "Valves Data".R13_XV06.MCMD,
                       fbk_open := "A/SSR_013_XV503_OFB",
                       fbk_close := "A/SSR_013_XV503_CFB",
                       reset := "Valves Data".R13_XV06.RESET OR "R13_DATA".R13.Reset,
                       intl := NOT "DI_INPUTS".R13_INPUTS_RUA.EMG_PB,
                       Mon_En := 1,
                       mon_sp := "Valves Data".R13_XV06.MON_TIME,
                       SEMI := "Valves Data".SEMI_AUTO.R13,
                       "open/close" => "A/SSR_013_XV503_CMD",
                       FAIL_TO_OPEN => "Valves Data".R13_VALVE_FAULT.XV06_FAIL_TO_OPEN,
                       FAIL_TO_CLOSE => "Valves Data".R13_VALVE_FAULT.XV06_FAIL_TO_CLOSE,
                       status => "Valves Data".R13_XV06.STATUS);
   END_IF;
END_REGION

REGION Network 138: R13_XV07
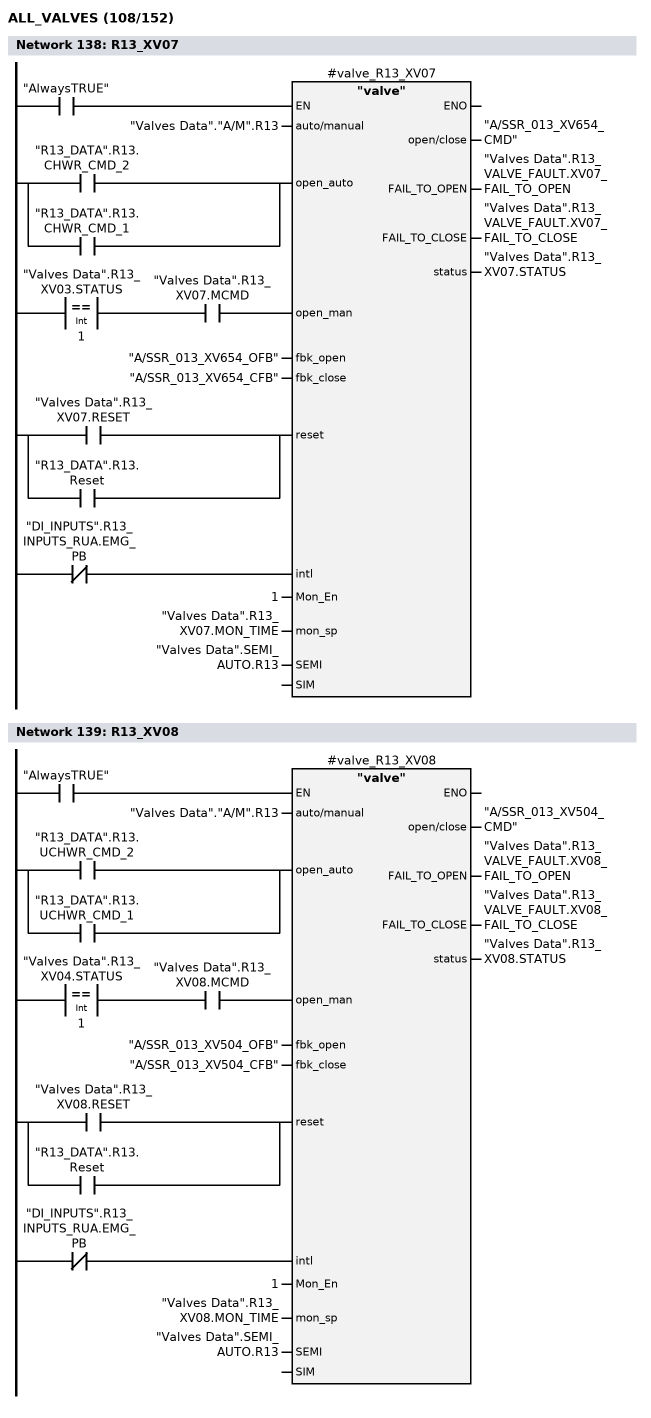
   RUNG wire#powerrail
      Contact( "AlwaysTRUE" )
      #valve_R13_XV07(open_auto := wire#w1, open_man := wire#w2, reset := wire#w3, intl := wire#w4, "auto/manual" := "Valves Data"."A/M".R13, fbk_open := "A/SSR_013_XV654_OFB", fbk_close := "A/SSR_013_XV654_CFB", Mon_En := 1, mon_sp := "Valves Data".R13_XV07.MON_TIME, SEMI := "Valves Data".SEMI_AUTO.R13, SIM :=, "open/close" => "A/SSR_013_XV654_CMD", FAIL_TO_OPEN => "Valves Data".R13_VALVE_FAULT.XV07_FAIL_TO_OPEN, FAIL_TO_CLOSE => "Valves Data".R13_VALVE_FAULT.XV07_FAIL_TO_CLOSE, status => "Valves Data".R13_XV07.STATUS)
   END_RUNG
   RUNG wire#powerrail
      Contact( "R13_DATA".R13.CHWR_CMD_2 )
   END_RUNG wire#w1
   RUNG wire#powerrail
      Contact( "R13_DATA".R13.CHWR_CMD_1 )
   END_RUNG wire#w1
   RUNG wire#powerrail
      { S7_Templates := "SrcType := Int" } EQ_Contact(in1 := "Valves Data".R13_XV03.STATUS, in2 := 1)
      Contact( "Valves Data".R13_XV07.MCMD )
   END_RUNG wire#w2
   RUNG wire#powerrail
      Contact( "Valves Data".R13_XV07.RESET )
   END_RUNG wire#w3
   RUNG wire#powerrail
      Contact( "R13_DATA".R13.Reset )
   END_RUNG wire#w3
   RUNG wire#powerrail
      I_Contact( "DI_INPUTS".R13_INPUTS_RUA.EMG_PB )
   END_RUNG wire#w4
   // the same network as SCL:
   IF "AlwaysTRUE" THEN
       #valve_R13_XV07("auto/manual" := "Valves Data"."A/M".R13,   // "valve"
                       open_auto := "R13_DATA".R13.CHWR_CMD_2 OR "R13_DATA".R13.CHWR_CMD_1,
                       open_man := ("Valves Data".R13_XV03.STATUS = 1) AND "Valves Data".R13_XV07.MCMD,
                       fbk_open := "A/SSR_013_XV654_OFB",
                       fbk_close := "A/SSR_013_XV654_CFB",
                       reset := "Valves Data".R13_XV07.RESET OR "R13_DATA".R13.Reset,
                       intl := NOT "DI_INPUTS".R13_INPUTS_RUA.EMG_PB,
                       Mon_En := 1,
                       mon_sp := "Valves Data".R13_XV07.MON_TIME,
                       SEMI := "Valves Data".SEMI_AUTO.R13,
                       "open/close" => "A/SSR_013_XV654_CMD",
                       FAIL_TO_OPEN => "Valves Data".R13_VALVE_FAULT.XV07_FAIL_TO_OPEN,
                       FAIL_TO_CLOSE => "Valves Data".R13_VALVE_FAULT.XV07_FAIL_TO_CLOSE,
                       status => "Valves Data".R13_XV07.STATUS);
   END_IF;
END_REGION

REGION Network 139: R13_XV08
   RUNG wire#powerrail
      Contact( "AlwaysTRUE" )
      #valve_R13_XV08(open_auto := wire#w1, open_man := wire#w2, reset := wire#w3, intl := wire#w4, "auto/manual" := "Valves Data"."A/M".R13, fbk_open := "A/SSR_013_XV504_OFB", fbk_close := "A/SSR_013_XV504_CFB", Mon_En := 1, mon_sp := "Valves Data".R13_XV08.MON_TIME, SEMI := "Valves Data".SEMI_AUTO.R13, SIM :=, "open/close" => "A/SSR_013_XV504_CMD", FAIL_TO_OPEN => "Valves Data".R13_VALVE_FAULT.XV08_FAIL_TO_OPEN, FAIL_TO_CLOSE => "Valves Data".R13_VALVE_FAULT.XV08_FAIL_TO_CLOSE, status => "Valves Data".R13_XV08.STATUS)
   END_RUNG
   RUNG wire#powerrail
      Contact( "R13_DATA".R13.UCHWR_CMD_2 )
   END_RUNG wire#w1
   RUNG wire#powerrail
      Contact( "R13_DATA".R13.UCHWR_CMD_1 )
   END_RUNG wire#w1
   RUNG wire#powerrail
      { S7_Templates := "SrcType := Int" } EQ_Contact(in1 := "Valves Data".R13_XV04.STATUS, in2 := 1)
      Contact( "Valves Data".R13_XV08.MCMD )
   END_RUNG wire#w2
   RUNG wire#powerrail
      Contact( "Valves Data".R13_XV08.RESET )
   END_RUNG wire#w3
   RUNG wire#powerrail
      Contact( "R13_DATA".R13.Reset )
   END_RUNG wire#w3
   RUNG wire#powerrail
      I_Contact( "DI_INPUTS".R13_INPUTS_RUA.EMG_PB )
   END_RUNG wire#w4
   // the same network as SCL:
   IF "AlwaysTRUE" THEN
       #valve_R13_XV08("auto/manual" := "Valves Data"."A/M".R13,   // "valve"
                       open_auto := "R13_DATA".R13.UCHWR_CMD_2 OR "R13_DATA".R13.UCHWR_CMD_1,
                       open_man := ("Valves Data".R13_XV04.STATUS = 1) AND "Valves Data".R13_XV08.MCMD,
                       fbk_open := "A/SSR_013_XV504_OFB",
                       fbk_close := "A/SSR_013_XV504_CFB",
                       reset := "Valves Data".R13_XV08.RESET OR "R13_DATA".R13.Reset,
                       intl := NOT "DI_INPUTS".R13_INPUTS_RUA.EMG_PB,
                       Mon_En := 1,
                       mon_sp := "Valves Data".R13_XV08.MON_TIME,
                       SEMI := "Valves Data".SEMI_AUTO.R13,
                       "open/close" => "A/SSR_013_XV504_CMD",
                       FAIL_TO_OPEN => "Valves Data".R13_VALVE_FAULT.XV08_FAIL_TO_OPEN,
                       FAIL_TO_CLOSE => "Valves Data".R13_VALVE_FAULT.XV08_FAIL_TO_CLOSE,
                       status => "Valves Data".R13_XV08.STATUS);
   END_IF;
END_REGION

REGION Network 140: R13_XV09
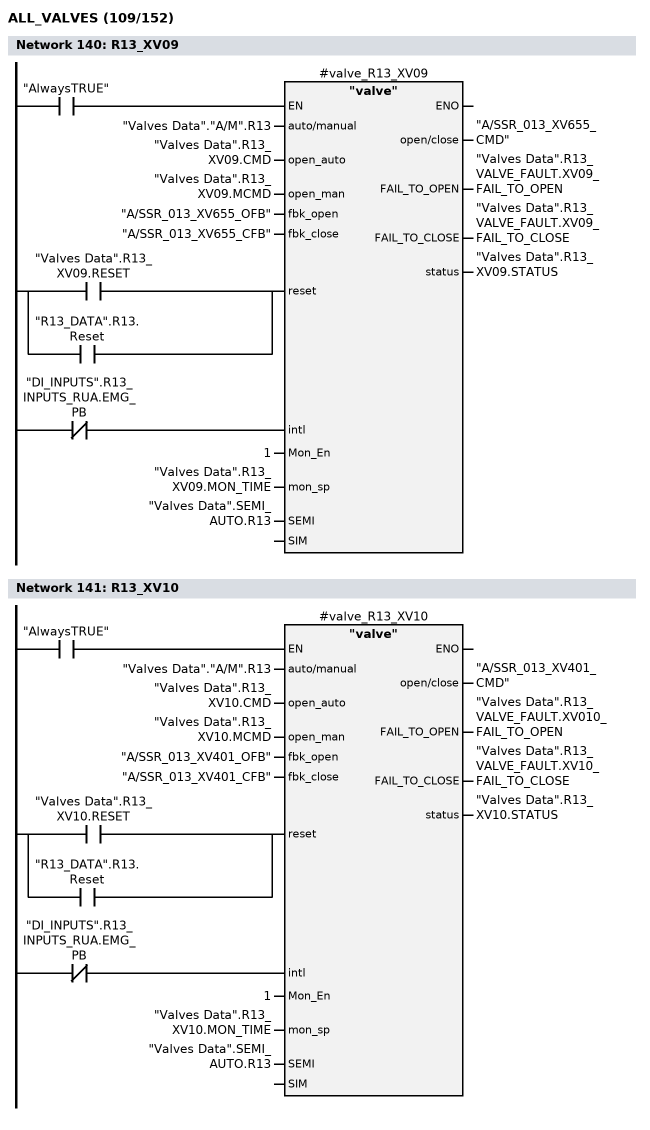
   RUNG wire#powerrail
      Contact( "AlwaysTRUE" )
      #valve_R13_XV09(reset := wire#w1, intl := wire#w2, "auto/manual" := "Valves Data"."A/M".R13, open_auto := "Valves Data".R13_XV09.CMD, open_man := "Valves Data".R13_XV09.MCMD, fbk_open := "A/SSR_013_XV655_OFB", fbk_close := "A/SSR_013_XV655_CFB", Mon_En := 1, mon_sp := "Valves Data".R13_XV09.MON_TIME, SEMI := "Valves Data".SEMI_AUTO.R13, SIM :=, "open/close" => "A/SSR_013_XV655_CMD", FAIL_TO_OPEN => "Valves Data".R13_VALVE_FAULT.XV09_FAIL_TO_OPEN, FAIL_TO_CLOSE => "Valves Data".R13_VALVE_FAULT.XV09_FAIL_TO_CLOSE, status => "Valves Data".R13_XV09.STATUS)
   END_RUNG
   RUNG wire#powerrail
      Contact( "Valves Data".R13_XV09.RESET )
   END_RUNG wire#w1
   RUNG wire#powerrail
      Contact( "R13_DATA".R13.Reset )
   END_RUNG wire#w1
   RUNG wire#powerrail
      I_Contact( "DI_INPUTS".R13_INPUTS_RUA.EMG_PB )
   END_RUNG wire#w2
   // the same network as SCL:
   IF "AlwaysTRUE" THEN
       #valve_R13_XV09("auto/manual" := "Valves Data"."A/M".R13,   // "valve"
                       open_auto := "Valves Data".R13_XV09.CMD,
                       open_man := "Valves Data".R13_XV09.MCMD,
                       fbk_open := "A/SSR_013_XV655_OFB",
                       fbk_close := "A/SSR_013_XV655_CFB",
                       reset := "Valves Data".R13_XV09.RESET OR "R13_DATA".R13.Reset,
                       intl := NOT "DI_INPUTS".R13_INPUTS_RUA.EMG_PB,
                       Mon_En := 1,
                       mon_sp := "Valves Data".R13_XV09.MON_TIME,
                       SEMI := "Valves Data".SEMI_AUTO.R13,
                       "open/close" => "A/SSR_013_XV655_CMD",
                       FAIL_TO_OPEN => "Valves Data".R13_VALVE_FAULT.XV09_FAIL_TO_OPEN,
                       FAIL_TO_CLOSE => "Valves Data".R13_VALVE_FAULT.XV09_FAIL_TO_CLOSE,
                       status => "Valves Data".R13_XV09.STATUS);
   END_IF;
END_REGION

REGION Network 141: R13_XV10
   RUNG wire#powerrail
      Contact( "AlwaysTRUE" )
      #valve_R13_XV10(reset := wire#w1, intl := wire#w2, "auto/manual" := "Valves Data"."A/M".R13, open_auto := "Valves Data".R13_XV10.CMD, open_man := "Valves Data".R13_XV10.MCMD, fbk_open := "A/SSR_013_XV401_OFB", fbk_close := "A/SSR_013_XV401_CFB", Mon_En := 1, mon_sp := "Valves Data".R13_XV10.MON_TIME, SEMI := "Valves Data".SEMI_AUTO.R13, SIM :=, "open/close" => "A/SSR_013_XV401_CMD", FAIL_TO_OPEN => "Valves Data".R13_VALVE_FAULT.XV010_FAIL_TO_OPEN, FAIL_TO_CLOSE => "Valves Data".R13_VALVE_FAULT.XV10_FAIL_TO_CLOSE, status => "Valves Data".R13_XV10.STATUS)
   END_RUNG
   RUNG wire#powerrail
      Contact( "Valves Data".R13_XV10.RESET )
   END_RUNG wire#w1
   RUNG wire#powerrail
      Contact( "R13_DATA".R13.Reset )
   END_RUNG wire#w1
   RUNG wire#powerrail
      I_Contact( "DI_INPUTS".R13_INPUTS_RUA.EMG_PB )
   END_RUNG wire#w2
   // the same network as SCL:
   IF "AlwaysTRUE" THEN
       #valve_R13_XV10("auto/manual" := "Valves Data"."A/M".R13,   // "valve"
                       open_auto := "Valves Data".R13_XV10.CMD,
                       open_man := "Valves Data".R13_XV10.MCMD,
                       fbk_open := "A/SSR_013_XV401_OFB",
                       fbk_close := "A/SSR_013_XV401_CFB",
                       reset := "Valves Data".R13_XV10.RESET OR "R13_DATA".R13.Reset,
                       intl := NOT "DI_INPUTS".R13_INPUTS_RUA.EMG_PB,
                       Mon_En := 1,
                       mon_sp := "Valves Data".R13_XV10.MON_TIME,
                       SEMI := "Valves Data".SEMI_AUTO.R13,
                       "open/close" => "A/SSR_013_XV401_CMD",
                       FAIL_TO_OPEN => "Valves Data".R13_VALVE_FAULT.XV010_FAIL_TO_OPEN,
                       FAIL_TO_CLOSE => "Valves Data".R13_VALVE_FAULT.XV10_FAIL_TO_CLOSE,
                       status => "Valves Data".R13_XV10.STATUS);
   END_IF;
END_REGION

REGION Network 142: ****REACTOR_14****
END_REGION

REGION Network 143: R14_XV01
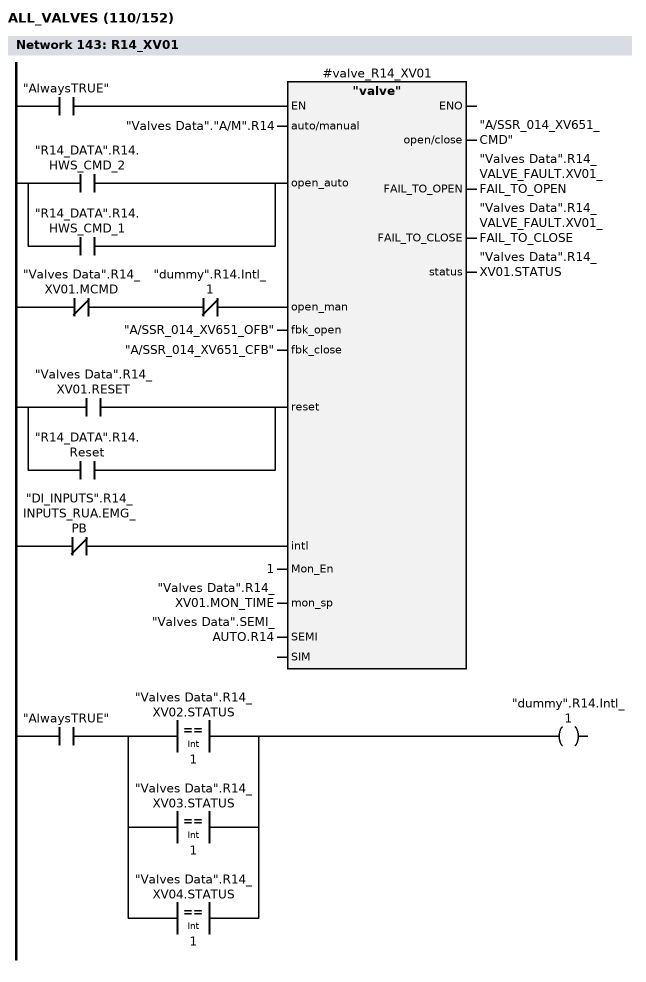
   RUNG wire#powerrail
      Contact( "AlwaysTRUE" )
      #valve_R14_XV01(open_auto := wire#w1, open_man := wire#w2, reset := wire#w3, intl := wire#w4, "auto/manual" := "Valves Data"."A/M".R14, fbk_open := "A/SSR_014_XV651_OFB", fbk_close := "A/SSR_014_XV651_CFB", Mon_En := 1, mon_sp := "Valves Data".R14_XV01.MON_TIME, SEMI := "Valves Data".SEMI_AUTO.R14, SIM :=, "open/close" => "A/SSR_014_XV651_CMD", FAIL_TO_OPEN => "Valves Data".R14_VALVE_FAULT.XV01_FAIL_TO_OPEN, FAIL_TO_CLOSE => "Valves Data".R14_VALVE_FAULT.XV01_FAIL_TO_CLOSE, status => "Valves Data".R14_XV01.STATUS)
   END_RUNG
   RUNG wire#powerrail
      Contact( "R14_DATA".R14.HWS_CMD_2 )
   END_RUNG wire#w1
   RUNG wire#powerrail
      Contact( "R14_DATA".R14.HWS_CMD_1 )
   END_RUNG wire#w1
   RUNG wire#powerrail
      I_Contact( "Valves Data".R14_XV01.MCMD )
      I_Contact( "dummy".R14.Intl_1 )
   END_RUNG wire#w2
   RUNG wire#powerrail
      Contact( "Valves Data".R14_XV01.RESET )
   END_RUNG wire#w3
   RUNG wire#powerrail
      Contact( "R14_DATA".R14.Reset )
   END_RUNG wire#w3
   RUNG wire#powerrail
      I_Contact( "DI_INPUTS".R14_INPUTS_RUA.EMG_PB )
   END_RUNG wire#w4
   RUNG wire#powerrail
      Contact( "AlwaysTRUE" )
      wire#w5
      { S7_Templates := "SrcType := Int" } EQ_Contact(in1 := "Valves Data".R14_XV02.STATUS, in2 := 1)
      wire#w6
      Coil( "dummy".R14.Intl_1 )
   END_RUNG
   RUNG wire#w5
      { S7_Templates := "SrcType := Int" } EQ_Contact(in1 := "Valves Data".R14_XV03.STATUS, in2 := 1)
   END_RUNG wire#w6
   RUNG wire#w5
      { S7_Templates := "SrcType := Int" } EQ_Contact(in1 := "Valves Data".R14_XV04.STATUS, in2 := 1)
   END_RUNG wire#w6
   // the same network as SCL:
   IF "AlwaysTRUE" THEN
       #valve_R14_XV01("auto/manual" := "Valves Data"."A/M".R14,   // "valve"
                       open_auto := "R14_DATA".R14.HWS_CMD_2 OR "R14_DATA".R14.HWS_CMD_1,
                       open_man := NOT "Valves Data".R14_XV01.MCMD AND NOT "dummy".R14.Intl_1,
                       fbk_open := "A/SSR_014_XV651_OFB",
                       fbk_close := "A/SSR_014_XV651_CFB",
                       reset := "Valves Data".R14_XV01.RESET OR "R14_DATA".R14.Reset,
                       intl := NOT "DI_INPUTS".R14_INPUTS_RUA.EMG_PB,
                       Mon_En := 1,
                       mon_sp := "Valves Data".R14_XV01.MON_TIME,
                       SEMI := "Valves Data".SEMI_AUTO.R14,
                       "open/close" => "A/SSR_014_XV651_CMD",
                       FAIL_TO_OPEN => "Valves Data".R14_VALVE_FAULT.XV01_FAIL_TO_OPEN,
                       FAIL_TO_CLOSE => "Valves Data".R14_VALVE_FAULT.XV01_FAIL_TO_CLOSE,
                       status => "Valves Data".R14_XV01.STATUS);
   END_IF;
   "dummy".R14.Intl_1 := "AlwaysTRUE" AND (("Valves Data".R14_XV02.STATUS = 1) OR ("Valves Data".R14_XV03.STATUS = 1) OR ("Valves Data".R14_XV04.STATUS = 1));
END_REGION

REGION Network 144: R14_XV02
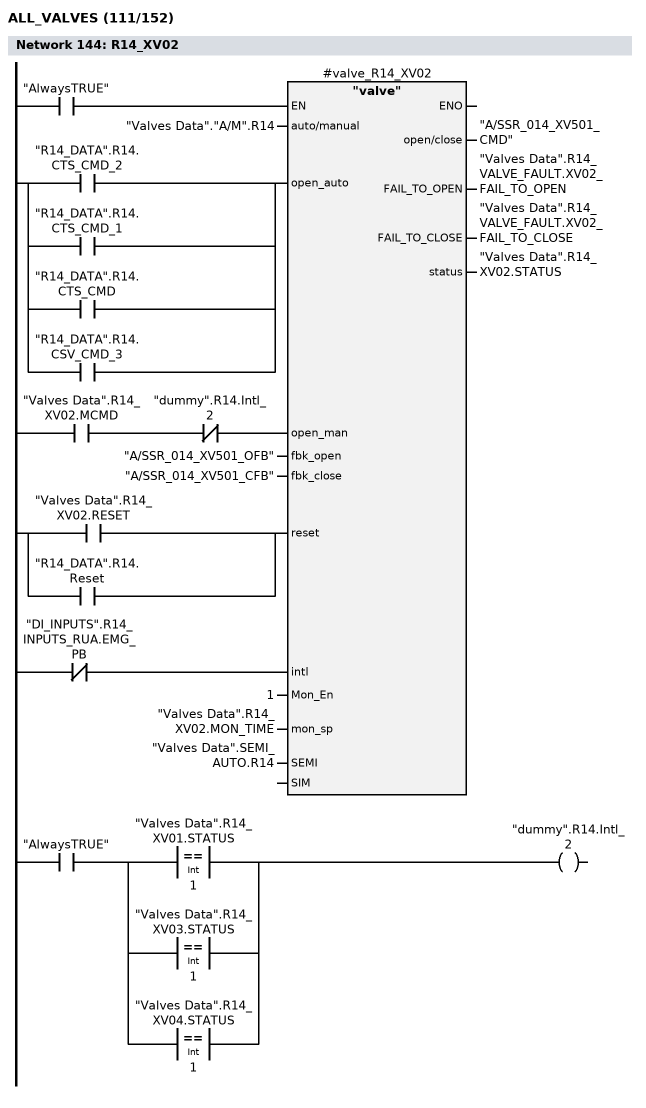
   RUNG wire#powerrail
      Contact( "AlwaysTRUE" )
      #valve_R14_XV02(open_auto := wire#w1, open_man := wire#w2, reset := wire#w3, intl := wire#w4, "auto/manual" := "Valves Data"."A/M".R14, fbk_open := "A/SSR_014_XV501_OFB", fbk_close := "A/SSR_014_XV501_CFB", Mon_En := 1, mon_sp := "Valves Data".R14_XV02.MON_TIME, SEMI := "Valves Data".SEMI_AUTO.R14, SIM :=, "open/close" => "A/SSR_014_XV501_CMD", FAIL_TO_OPEN => "Valves Data".R14_VALVE_FAULT.XV02_FAIL_TO_OPEN, FAIL_TO_CLOSE => "Valves Data".R14_VALVE_FAULT.XV02_FAIL_TO_CLOSE, status => "Valves Data".R14_XV02.STATUS)
   END_RUNG
   RUNG wire#powerrail
      Contact( "R14_DATA".R14.CTS_CMD_2 )
   END_RUNG wire#w1
   RUNG wire#powerrail
      Contact( "R14_DATA".R14.CTS_CMD_1 )
   END_RUNG wire#w1
   RUNG wire#powerrail
      Contact( "R14_DATA".R14.CTS_CMD )
   END_RUNG wire#w1
   RUNG wire#powerrail
      Contact( "R14_DATA".R14.CSV_CMD_3 )
   END_RUNG wire#w1
   RUNG wire#powerrail
      Contact( "Valves Data".R14_XV02.MCMD )
      I_Contact( "dummy".R14.Intl_2 )
   END_RUNG wire#w2
   RUNG wire#powerrail
      Contact( "Valves Data".R14_XV02.RESET )
   END_RUNG wire#w3
   RUNG wire#powerrail
      Contact( "R14_DATA".R14.Reset )
   END_RUNG wire#w3
   RUNG wire#powerrail
      I_Contact( "DI_INPUTS".R14_INPUTS_RUA.EMG_PB )
   END_RUNG wire#w4
   RUNG wire#powerrail
      Contact( "AlwaysTRUE" )
      wire#w5
      { S7_Templates := "SrcType := Int" } EQ_Contact(in1 := "Valves Data".R14_XV01.STATUS, in2 := 1)
      wire#w6
      Coil( "dummy".R14.Intl_2 )
   END_RUNG
   RUNG wire#w5
      { S7_Templates := "SrcType := Int" } EQ_Contact(in1 := "Valves Data".R14_XV03.STATUS, in2 := 1)
   END_RUNG wire#w6
   RUNG wire#w5
      { S7_Templates := "SrcType := Int" } EQ_Contact(in1 := "Valves Data".R14_XV04.STATUS, in2 := 1)
   END_RUNG wire#w6
   // the same network as SCL:
   IF "AlwaysTRUE" THEN
       #valve_R14_XV02("auto/manual" := "Valves Data"."A/M".R14,   // "valve"
                       open_auto := "R14_DATA".R14.CTS_CMD_2 OR "R14_DATA".R14.CTS_CMD_1 OR "R14_DATA".R14.CTS_CMD OR "R14_DATA".R14.CSV_CMD_3,
                       open_man := "Valves Data".R14_XV02.MCMD AND NOT "dummy".R14.Intl_2,
                       fbk_open := "A/SSR_014_XV501_OFB",
                       fbk_close := "A/SSR_014_XV501_CFB",
                       reset := "Valves Data".R14_XV02.RESET OR "R14_DATA".R14.Reset,
                       intl := NOT "DI_INPUTS".R14_INPUTS_RUA.EMG_PB,
                       Mon_En := 1,
                       mon_sp := "Valves Data".R14_XV02.MON_TIME,
                       SEMI := "Valves Data".SEMI_AUTO.R14,
                       "open/close" => "A/SSR_014_XV501_CMD",
                       FAIL_TO_OPEN => "Valves Data".R14_VALVE_FAULT.XV02_FAIL_TO_OPEN,
                       FAIL_TO_CLOSE => "Valves Data".R14_VALVE_FAULT.XV02_FAIL_TO_CLOSE,
                       status => "Valves Data".R14_XV02.STATUS);
   END_IF;
   "dummy".R14.Intl_2 := "AlwaysTRUE" AND (("Valves Data".R14_XV01.STATUS = 1) OR ("Valves Data".R14_XV03.STATUS = 1) OR ("Valves Data".R14_XV04.STATUS = 1));
END_REGION

REGION Network 145: R14_XV03
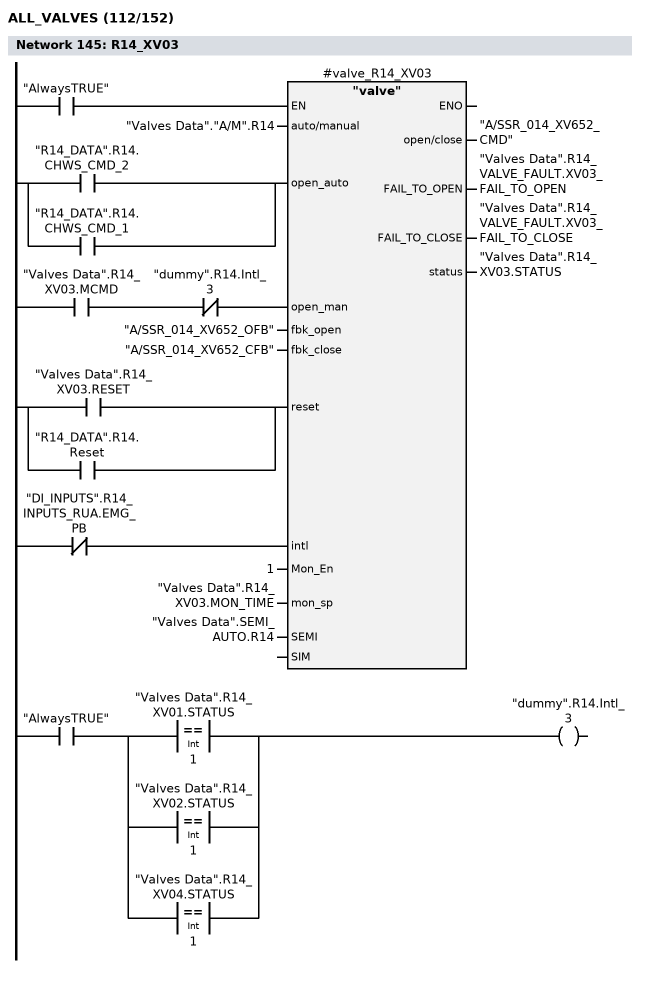
   RUNG wire#powerrail
      Contact( "AlwaysTRUE" )
      #valve_R14_XV03(open_auto := wire#w1, open_man := wire#w2, reset := wire#w3, intl := wire#w4, "auto/manual" := "Valves Data"."A/M".R14, fbk_open := "A/SSR_014_XV652_OFB", fbk_close := "A/SSR_014_XV652_CFB", Mon_En := 1, mon_sp := "Valves Data".R14_XV03.MON_TIME, SEMI := "Valves Data".SEMI_AUTO.R14, SIM :=, "open/close" => "A/SSR_014_XV652_CMD", FAIL_TO_OPEN => "Valves Data".R14_VALVE_FAULT.XV03_FAIL_TO_OPEN, FAIL_TO_CLOSE => "Valves Data".R14_VALVE_FAULT.XV03_FAIL_TO_CLOSE, status => "Valves Data".R14_XV03.STATUS)
   END_RUNG
   RUNG wire#powerrail
      Contact( "R14_DATA".R14.CHWS_CMD_2 )
   END_RUNG wire#w1
   RUNG wire#powerrail
      Contact( "R14_DATA".R14.CHWS_CMD_1 )
   END_RUNG wire#w1
   RUNG wire#powerrail
      Contact( "Valves Data".R14_XV03.MCMD )
      I_Contact( "dummy".R14.Intl_3 )
   END_RUNG wire#w2
   RUNG wire#powerrail
      Contact( "Valves Data".R14_XV03.RESET )
   END_RUNG wire#w3
   RUNG wire#powerrail
      Contact( "R14_DATA".R14.Reset )
   END_RUNG wire#w3
   RUNG wire#powerrail
      I_Contact( "DI_INPUTS".R14_INPUTS_RUA.EMG_PB )
   END_RUNG wire#w4
   RUNG wire#powerrail
      Contact( "AlwaysTRUE" )
      wire#w5
      { S7_Templates := "SrcType := Int" } EQ_Contact(in1 := "Valves Data".R14_XV01.STATUS, in2 := 1)
      wire#w6
      Coil( "dummy".R14.Intl_3 )
   END_RUNG
   RUNG wire#w5
      { S7_Templates := "SrcType := Int" } EQ_Contact(in1 := "Valves Data".R14_XV02.STATUS, in2 := 1)
   END_RUNG wire#w6
   RUNG wire#w5
      { S7_Templates := "SrcType := Int" } EQ_Contact(in1 := "Valves Data".R14_XV04.STATUS, in2 := 1)
   END_RUNG wire#w6
   // the same network as SCL:
   IF "AlwaysTRUE" THEN
       #valve_R14_XV03("auto/manual" := "Valves Data"."A/M".R14,   // "valve"
                       open_auto := "R14_DATA".R14.CHWS_CMD_2 OR "R14_DATA".R14.CHWS_CMD_1,
                       open_man := "Valves Data".R14_XV03.MCMD AND NOT "dummy".R14.Intl_3,
                       fbk_open := "A/SSR_014_XV652_OFB",
                       fbk_close := "A/SSR_014_XV652_CFB",
                       reset := "Valves Data".R14_XV03.RESET OR "R14_DATA".R14.Reset,
                       intl := NOT "DI_INPUTS".R14_INPUTS_RUA.EMG_PB,
                       Mon_En := 1,
                       mon_sp := "Valves Data".R14_XV03.MON_TIME,
                       SEMI := "Valves Data".SEMI_AUTO.R14,
                       "open/close" => "A/SSR_014_XV652_CMD",
                       FAIL_TO_OPEN => "Valves Data".R14_VALVE_FAULT.XV03_FAIL_TO_OPEN,
                       FAIL_TO_CLOSE => "Valves Data".R14_VALVE_FAULT.XV03_FAIL_TO_CLOSE,
                       status => "Valves Data".R14_XV03.STATUS);
   END_IF;
   "dummy".R14.Intl_3 := "AlwaysTRUE" AND (("Valves Data".R14_XV01.STATUS = 1) OR ("Valves Data".R14_XV02.STATUS = 1) OR ("Valves Data".R14_XV04.STATUS = 1));
END_REGION

REGION Network 146: R14_XV04
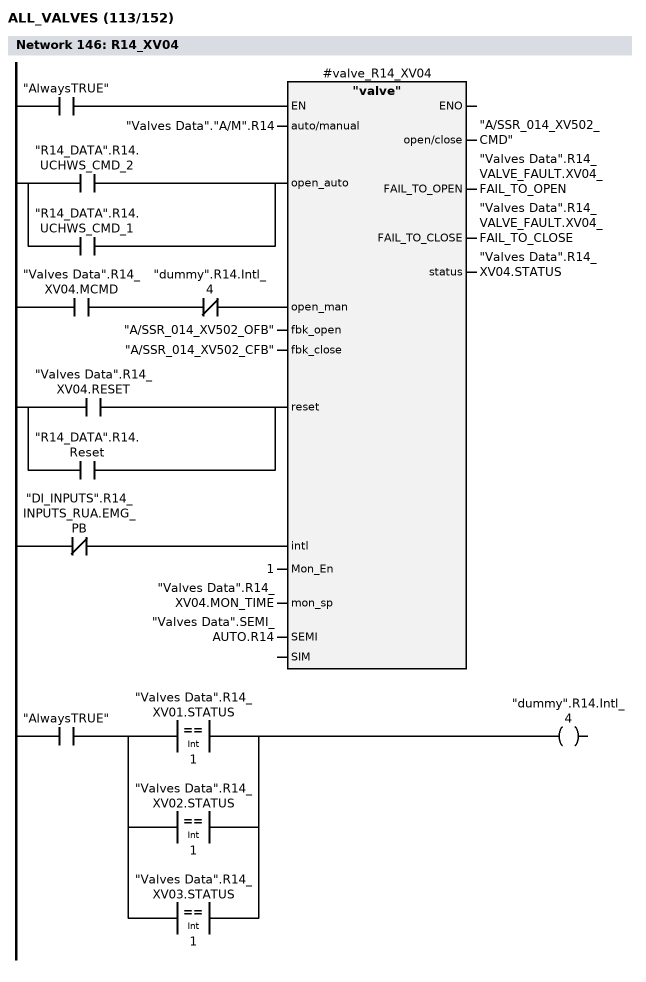
   RUNG wire#powerrail
      Contact( "AlwaysTRUE" )
      #valve_R14_XV04(open_auto := wire#w1, open_man := wire#w2, reset := wire#w3, intl := wire#w4, "auto/manual" := "Valves Data"."A/M".R14, fbk_open := "A/SSR_014_XV502_OFB", fbk_close := "A/SSR_014_XV502_CFB", Mon_En := 1, mon_sp := "Valves Data".R14_XV04.MON_TIME, SEMI := "Valves Data".SEMI_AUTO.R14, SIM :=, "open/close" => "A/SSR_014_XV502_CMD", FAIL_TO_OPEN => "Valves Data".R14_VALVE_FAULT.XV04_FAIL_TO_OPEN, FAIL_TO_CLOSE => "Valves Data".R14_VALVE_FAULT.XV04_FAIL_TO_CLOSE, status => "Valves Data".R14_XV04.STATUS)
   END_RUNG
   RUNG wire#powerrail
      Contact( "R14_DATA".R14.UCHWS_CMD_2 )
   END_RUNG wire#w1
   RUNG wire#powerrail
      Contact( "R14_DATA".R14.UCHWS_CMD_1 )
   END_RUNG wire#w1
   RUNG wire#powerrail
      Contact( "Valves Data".R14_XV04.MCMD )
      I_Contact( "dummy".R14.Intl_4 )
   END_RUNG wire#w2
   RUNG wire#powerrail
      Contact( "Valves Data".R14_XV04.RESET )
   END_RUNG wire#w3
   RUNG wire#powerrail
      Contact( "R14_DATA".R14.Reset )
   END_RUNG wire#w3
   RUNG wire#powerrail
      I_Contact( "DI_INPUTS".R14_INPUTS_RUA.EMG_PB )
   END_RUNG wire#w4
   RUNG wire#powerrail
      Contact( "AlwaysTRUE" )
      wire#w5
      { S7_Templates := "SrcType := Int" } EQ_Contact(in1 := "Valves Data".R14_XV01.STATUS, in2 := 1)
      wire#w6
      Coil( "dummy".R14.Intl_4 )
   END_RUNG
   RUNG wire#w5
      { S7_Templates := "SrcType := Int" } EQ_Contact(in1 := "Valves Data".R14_XV02.STATUS, in2 := 1)
   END_RUNG wire#w6
   RUNG wire#w5
      { S7_Templates := "SrcType := Int" } EQ_Contact(in1 := "Valves Data".R14_XV03.STATUS, in2 := 1)
   END_RUNG wire#w6
   // the same network as SCL:
   IF "AlwaysTRUE" THEN
       #valve_R14_XV04("auto/manual" := "Valves Data"."A/M".R14,   // "valve"
                       open_auto := "R14_DATA".R14.UCHWS_CMD_2 OR "R14_DATA".R14.UCHWS_CMD_1,
                       open_man := "Valves Data".R14_XV04.MCMD AND NOT "dummy".R14.Intl_4,
                       fbk_open := "A/SSR_014_XV502_OFB",
                       fbk_close := "A/SSR_014_XV502_CFB",
                       reset := "Valves Data".R14_XV04.RESET OR "R14_DATA".R14.Reset,
                       intl := NOT "DI_INPUTS".R14_INPUTS_RUA.EMG_PB,
                       Mon_En := 1,
                       mon_sp := "Valves Data".R14_XV04.MON_TIME,
                       SEMI := "Valves Data".SEMI_AUTO.R14,
                       "open/close" => "A/SSR_014_XV502_CMD",
                       FAIL_TO_OPEN => "Valves Data".R14_VALVE_FAULT.XV04_FAIL_TO_OPEN,
                       FAIL_TO_CLOSE => "Valves Data".R14_VALVE_FAULT.XV04_FAIL_TO_CLOSE,
                       status => "Valves Data".R14_XV04.STATUS);
   END_IF;
   "dummy".R14.Intl_4 := "AlwaysTRUE" AND (("Valves Data".R14_XV01.STATUS = 1) OR ("Valves Data".R14_XV02.STATUS = 1) OR ("Valves Data".R14_XV03.STATUS = 1));
END_REGION

REGION Network 147: R14_XV05
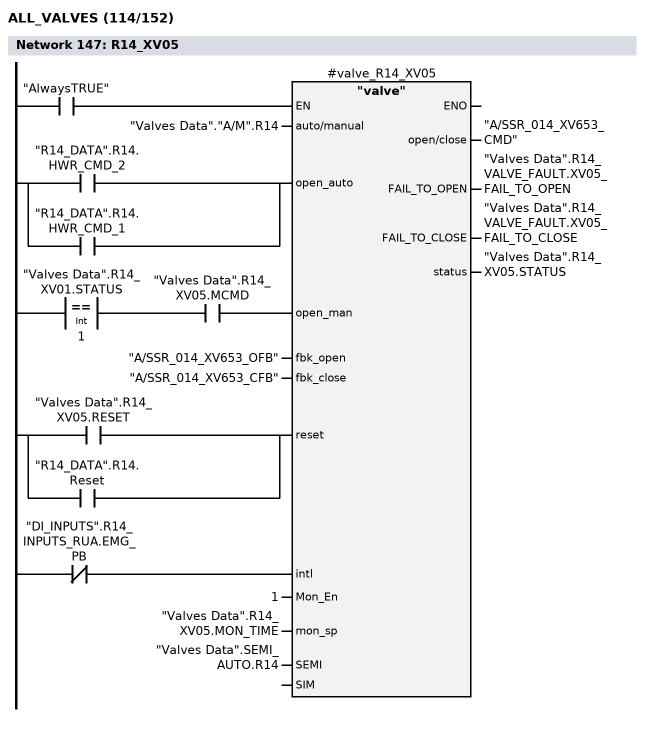
   RUNG wire#powerrail
      Contact( "AlwaysTRUE" )
      #valve_R14_XV05(open_auto := wire#w1, open_man := wire#w2, reset := wire#w3, intl := wire#w4, "auto/manual" := "Valves Data"."A/M".R14, fbk_open := "A/SSR_014_XV653_OFB", fbk_close := "A/SSR_014_XV653_CFB", Mon_En := 1, mon_sp := "Valves Data".R14_XV05.MON_TIME, SEMI := "Valves Data".SEMI_AUTO.R14, SIM :=, "open/close" => "A/SSR_014_XV653_CMD", FAIL_TO_OPEN => "Valves Data".R14_VALVE_FAULT.XV05_FAIL_TO_OPEN, FAIL_TO_CLOSE => "Valves Data".R14_VALVE_FAULT.XV05_FAIL_TO_CLOSE, status => "Valves Data".R14_XV05.STATUS)
   END_RUNG
   RUNG wire#powerrail
      Contact( "R14_DATA".R14.HWR_CMD_2 )
   END_RUNG wire#w1
   RUNG wire#powerrail
      Contact( "R14_DATA".R14.HWR_CMD_1 )
   END_RUNG wire#w1
   RUNG wire#powerrail
      { S7_Templates := "SrcType := Int" } EQ_Contact(in1 := "Valves Data".R14_XV01.STATUS, in2 := 1)
      Contact( "Valves Data".R14_XV05.MCMD )
   END_RUNG wire#w2
   RUNG wire#powerrail
      Contact( "Valves Data".R14_XV05.RESET )
   END_RUNG wire#w3
   RUNG wire#powerrail
      Contact( "R14_DATA".R14.Reset )
   END_RUNG wire#w3
   RUNG wire#powerrail
      I_Contact( "DI_INPUTS".R14_INPUTS_RUA.EMG_PB )
   END_RUNG wire#w4
   // the same network as SCL:
   IF "AlwaysTRUE" THEN
       #valve_R14_XV05("auto/manual" := "Valves Data"."A/M".R14,   // "valve"
                       open_auto := "R14_DATA".R14.HWR_CMD_2 OR "R14_DATA".R14.HWR_CMD_1,
                       open_man := ("Valves Data".R14_XV01.STATUS = 1) AND "Valves Data".R14_XV05.MCMD,
                       fbk_open := "A/SSR_014_XV653_OFB",
                       fbk_close := "A/SSR_014_XV653_CFB",
                       reset := "Valves Data".R14_XV05.RESET OR "R14_DATA".R14.Reset,
                       intl := NOT "DI_INPUTS".R14_INPUTS_RUA.EMG_PB,
                       Mon_En := 1,
                       mon_sp := "Valves Data".R14_XV05.MON_TIME,
                       SEMI := "Valves Data".SEMI_AUTO.R14,
                       "open/close" => "A/SSR_014_XV653_CMD",
                       FAIL_TO_OPEN => "Valves Data".R14_VALVE_FAULT.XV05_FAIL_TO_OPEN,
                       FAIL_TO_CLOSE => "Valves Data".R14_VALVE_FAULT.XV05_FAIL_TO_CLOSE,
                       status => "Valves Data".R14_XV05.STATUS);
   END_IF;
END_REGION

REGION Network 148: R14_XV06
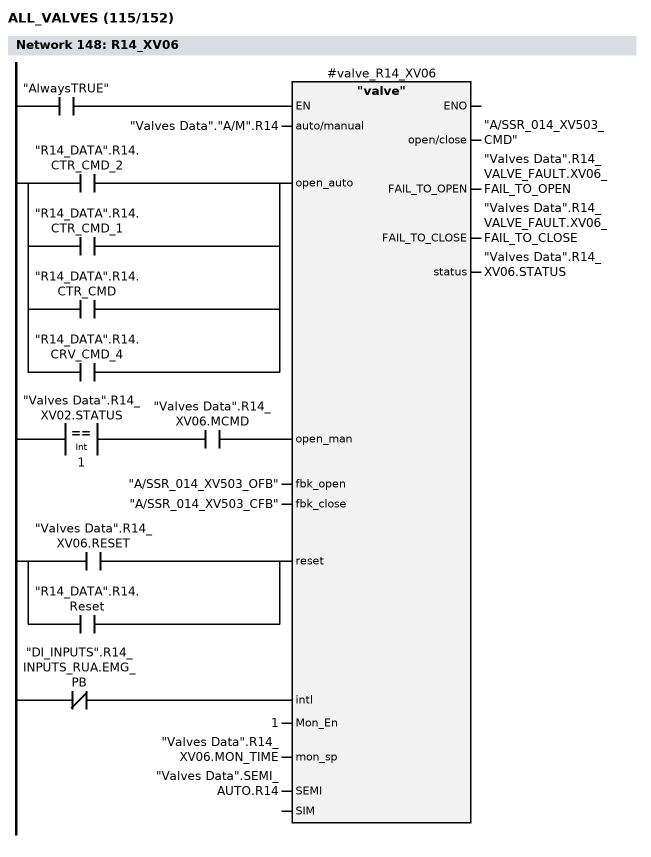
   RUNG wire#powerrail
      Contact( "AlwaysTRUE" )
      #valve_R14_XV06(open_auto := wire#w1, open_man := wire#w2, reset := wire#w3, intl := wire#w4, "auto/manual" := "Valves Data"."A/M".R14, fbk_open := "A/SSR_014_XV503_OFB", fbk_close := "A/SSR_014_XV503_CFB", Mon_En := 1, mon_sp := "Valves Data".R14_XV06.MON_TIME, SEMI := "Valves Data".SEMI_AUTO.R14, SIM :=, "open/close" => "A/SSR_014_XV503_CMD", FAIL_TO_OPEN => "Valves Data".R14_VALVE_FAULT.XV06_FAIL_TO_OPEN, FAIL_TO_CLOSE => "Valves Data".R14_VALVE_FAULT.XV06_FAIL_TO_CLOSE, status => "Valves Data".R14_XV06.STATUS)
   END_RUNG
   RUNG wire#powerrail
      Contact( "R14_DATA".R14.CTR_CMD_2 )
   END_RUNG wire#w1
   RUNG wire#powerrail
      Contact( "R14_DATA".R14.CTR_CMD_1 )
   END_RUNG wire#w1
   RUNG wire#powerrail
      Contact( "R14_DATA".R14.CTR_CMD )
   END_RUNG wire#w1
   RUNG wire#powerrail
      Contact( "R14_DATA".R14.CRV_CMD_4 )
   END_RUNG wire#w1
   RUNG wire#powerrail
      { S7_Templates := "SrcType := Int" } EQ_Contact(in1 := "Valves Data".R14_XV02.STATUS, in2 := 1)
      Contact( "Valves Data".R14_XV06.MCMD )
   END_RUNG wire#w2
   RUNG wire#powerrail
      Contact( "Valves Data".R14_XV06.RESET )
   END_RUNG wire#w3
   RUNG wire#powerrail
      Contact( "R14_DATA".R14.Reset )
   END_RUNG wire#w3
   RUNG wire#powerrail
      I_Contact( "DI_INPUTS".R14_INPUTS_RUA.EMG_PB )
   END_RUNG wire#w4
   // the same network as SCL:
   IF "AlwaysTRUE" THEN
       #valve_R14_XV06("auto/manual" := "Valves Data"."A/M".R14,   // "valve"
                       open_auto := "R14_DATA".R14.CTR_CMD_2 OR "R14_DATA".R14.CTR_CMD_1 OR "R14_DATA".R14.CTR_CMD OR "R14_DATA".R14.CRV_CMD_4,
                       open_man := ("Valves Data".R14_XV02.STATUS = 1) AND "Valves Data".R14_XV06.MCMD,
                       fbk_open := "A/SSR_014_XV503_OFB",
                       fbk_close := "A/SSR_014_XV503_CFB",
                       reset := "Valves Data".R14_XV06.RESET OR "R14_DATA".R14.Reset,
                       intl := NOT "DI_INPUTS".R14_INPUTS_RUA.EMG_PB,
                       Mon_En := 1,
                       mon_sp := "Valves Data".R14_XV06.MON_TIME,
                       SEMI := "Valves Data".SEMI_AUTO.R14,
                       "open/close" => "A/SSR_014_XV503_CMD",
                       FAIL_TO_OPEN => "Valves Data".R14_VALVE_FAULT.XV06_FAIL_TO_OPEN,
                       FAIL_TO_CLOSE => "Valves Data".R14_VALVE_FAULT.XV06_FAIL_TO_CLOSE,
                       status => "Valves Data".R14_XV06.STATUS);
   END_IF;
END_REGION

REGION Network 149: R14_XV07
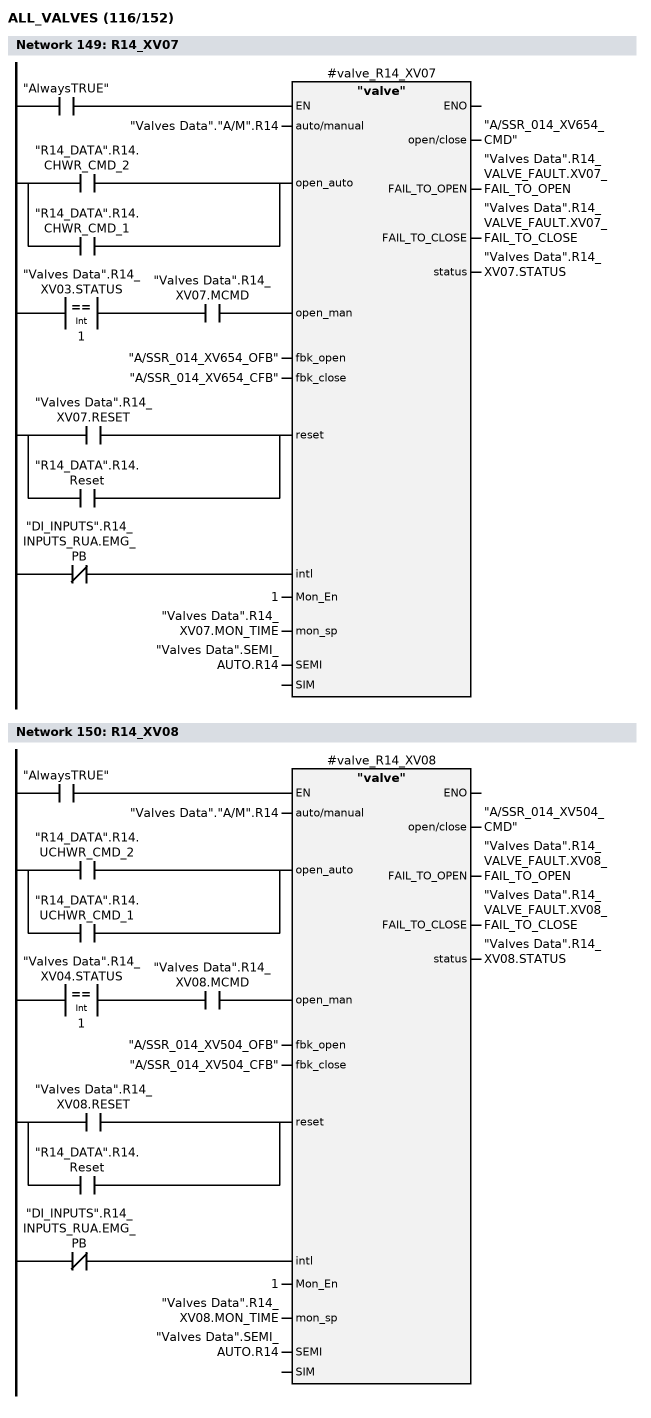
   RUNG wire#powerrail
      Contact( "AlwaysTRUE" )
      #valve_R14_XV07(open_auto := wire#w1, open_man := wire#w2, reset := wire#w3, intl := wire#w4, "auto/manual" := "Valves Data"."A/M".R14, fbk_open := "A/SSR_014_XV654_OFB", fbk_close := "A/SSR_014_XV654_CFB", Mon_En := 1, mon_sp := "Valves Data".R14_XV07.MON_TIME, SEMI := "Valves Data".SEMI_AUTO.R14, SIM :=, "open/close" => "A/SSR_014_XV654_CMD", FAIL_TO_OPEN => "Valves Data".R14_VALVE_FAULT.XV07_FAIL_TO_OPEN, FAIL_TO_CLOSE => "Valves Data".R14_VALVE_FAULT.XV07_FAIL_TO_CLOSE, status => "Valves Data".R14_XV07.STATUS)
   END_RUNG
   RUNG wire#powerrail
      Contact( "R14_DATA".R14.CHWR_CMD_2 )
   END_RUNG wire#w1
   RUNG wire#powerrail
      Contact( "R14_DATA".R14.CHWR_CMD_1 )
   END_RUNG wire#w1
   RUNG wire#powerrail
      { S7_Templates := "SrcType := Int" } EQ_Contact(in1 := "Valves Data".R14_XV03.STATUS, in2 := 1)
      Contact( "Valves Data".R14_XV07.MCMD )
   END_RUNG wire#w2
   RUNG wire#powerrail
      Contact( "Valves Data".R14_XV07.RESET )
   END_RUNG wire#w3
   RUNG wire#powerrail
      Contact( "R14_DATA".R14.Reset )
   END_RUNG wire#w3
   RUNG wire#powerrail
      I_Contact( "DI_INPUTS".R14_INPUTS_RUA.EMG_PB )
   END_RUNG wire#w4
   // the same network as SCL:
   IF "AlwaysTRUE" THEN
       #valve_R14_XV07("auto/manual" := "Valves Data"."A/M".R14,   // "valve"
                       open_auto := "R14_DATA".R14.CHWR_CMD_2 OR "R14_DATA".R14.CHWR_CMD_1,
                       open_man := ("Valves Data".R14_XV03.STATUS = 1) AND "Valves Data".R14_XV07.MCMD,
                       fbk_open := "A/SSR_014_XV654_OFB",
                       fbk_close := "A/SSR_014_XV654_CFB",
                       reset := "Valves Data".R14_XV07.RESET OR "R14_DATA".R14.Reset,
                       intl := NOT "DI_INPUTS".R14_INPUTS_RUA.EMG_PB,
                       Mon_En := 1,
                       mon_sp := "Valves Data".R14_XV07.MON_TIME,
                       SEMI := "Valves Data".SEMI_AUTO.R14,
                       "open/close" => "A/SSR_014_XV654_CMD",
                       FAIL_TO_OPEN => "Valves Data".R14_VALVE_FAULT.XV07_FAIL_TO_OPEN,
                       FAIL_TO_CLOSE => "Valves Data".R14_VALVE_FAULT.XV07_FAIL_TO_CLOSE,
                       status => "Valves Data".R14_XV07.STATUS);
   END_IF;
END_REGION

REGION Network 150: R14_XV08
   RUNG wire#powerrail
      Contact( "AlwaysTRUE" )
      #valve_R14_XV08(open_auto := wire#w1, open_man := wire#w2, reset := wire#w3, intl := wire#w4, "auto/manual" := "Valves Data"."A/M".R14, fbk_open := "A/SSR_014_XV504_OFB", fbk_close := "A/SSR_014_XV504_CFB", Mon_En := 1, mon_sp := "Valves Data".R14_XV08.MON_TIME, SEMI := "Valves Data".SEMI_AUTO.R14, SIM :=, "open/close" => "A/SSR_014_XV504_CMD", FAIL_TO_OPEN => "Valves Data".R14_VALVE_FAULT.XV08_FAIL_TO_OPEN, FAIL_TO_CLOSE => "Valves Data".R14_VALVE_FAULT.XV08_FAIL_TO_CLOSE, status => "Valves Data".R14_XV08.STATUS)
   END_RUNG
   RUNG wire#powerrail
      Contact( "R14_DATA".R14.UCHWR_CMD_2 )
   END_RUNG wire#w1
   RUNG wire#powerrail
      Contact( "R14_DATA".R14.UCHWR_CMD_1 )
   END_RUNG wire#w1
   RUNG wire#powerrail
      { S7_Templates := "SrcType := Int" } EQ_Contact(in1 := "Valves Data".R14_XV04.STATUS, in2 := 1)
      Contact( "Valves Data".R14_XV08.MCMD )
   END_RUNG wire#w2
   RUNG wire#powerrail
      Contact( "Valves Data".R14_XV08.RESET )
   END_RUNG wire#w3
   RUNG wire#powerrail
      Contact( "R14_DATA".R14.Reset )
   END_RUNG wire#w3
   RUNG wire#powerrail
      I_Contact( "DI_INPUTS".R14_INPUTS_RUA.EMG_PB )
   END_RUNG wire#w4
   // the same network as SCL:
   IF "AlwaysTRUE" THEN
       #valve_R14_XV08("auto/manual" := "Valves Data"."A/M".R14,   // "valve"
                       open_auto := "R14_DATA".R14.UCHWR_CMD_2 OR "R14_DATA".R14.UCHWR_CMD_1,
                       open_man := ("Valves Data".R14_XV04.STATUS = 1) AND "Valves Data".R14_XV08.MCMD,
                       fbk_open := "A/SSR_014_XV504_OFB",
                       fbk_close := "A/SSR_014_XV504_CFB",
                       reset := "Valves Data".R14_XV08.RESET OR "R14_DATA".R14.Reset,
                       intl := NOT "DI_INPUTS".R14_INPUTS_RUA.EMG_PB,
                       Mon_En := 1,
                       mon_sp := "Valves Data".R14_XV08.MON_TIME,
                       SEMI := "Valves Data".SEMI_AUTO.R14,
                       "open/close" => "A/SSR_014_XV504_CMD",
                       FAIL_TO_OPEN => "Valves Data".R14_VALVE_FAULT.XV08_FAIL_TO_OPEN,
                       FAIL_TO_CLOSE => "Valves Data".R14_VALVE_FAULT.XV08_FAIL_TO_CLOSE,
                       status => "Valves Data".R14_XV08.STATUS);
   END_IF;
END_REGION

REGION Network 151: R14_XV09
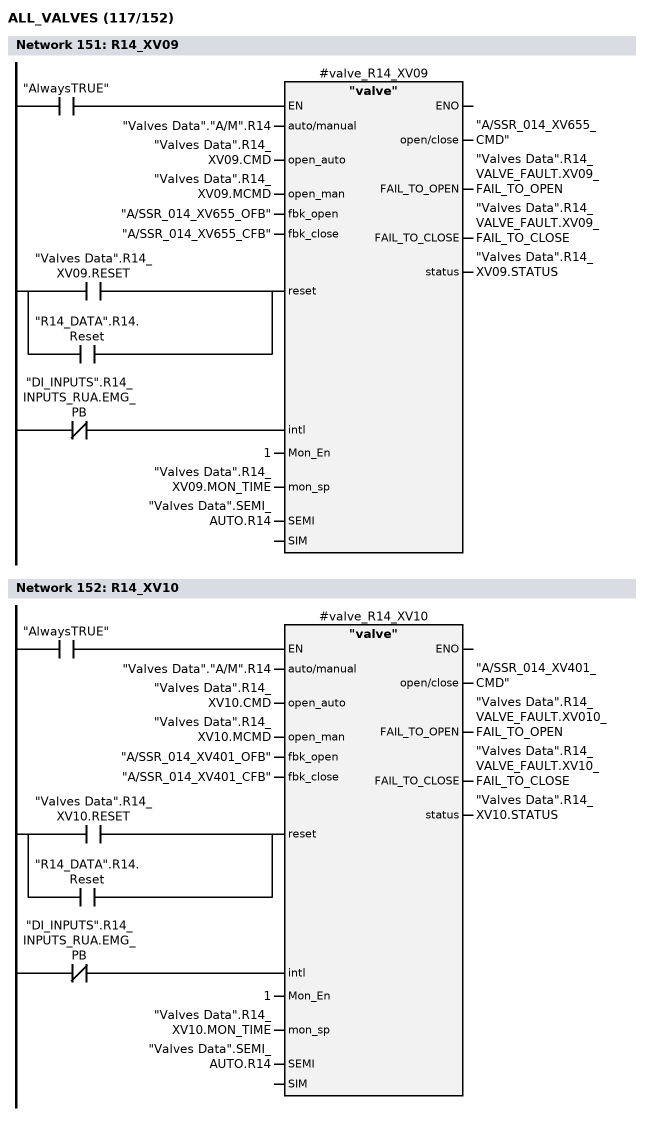
   RUNG wire#powerrail
      Contact( "AlwaysTRUE" )
      #valve_R14_XV09(reset := wire#w1, intl := wire#w2, "auto/manual" := "Valves Data"."A/M".R14, open_auto := "Valves Data".R14_XV09.CMD, open_man := "Valves Data".R14_XV09.MCMD, fbk_open := "A/SSR_014_XV655_OFB", fbk_close := "A/SSR_014_XV655_CFB", Mon_En := 1, mon_sp := "Valves Data".R14_XV09.MON_TIME, SEMI := "Valves Data".SEMI_AUTO.R14, SIM :=, "open/close" => "A/SSR_014_XV655_CMD", FAIL_TO_OPEN => "Valves Data".R14_VALVE_FAULT.XV09_FAIL_TO_OPEN, FAIL_TO_CLOSE => "Valves Data".R14_VALVE_FAULT.XV09_FAIL_TO_CLOSE, status => "Valves Data".R14_XV09.STATUS)
   END_RUNG
   RUNG wire#powerrail
      Contact( "Valves Data".R14_XV09.RESET )
   END_RUNG wire#w1
   RUNG wire#powerrail
      Contact( "R14_DATA".R14.Reset )
   END_RUNG wire#w1
   RUNG wire#powerrail
      I_Contact( "DI_INPUTS".R14_INPUTS_RUA.EMG_PB )
   END_RUNG wire#w2
   // the same network as SCL:
   IF "AlwaysTRUE" THEN
       #valve_R14_XV09("auto/manual" := "Valves Data"."A/M".R14,   // "valve"
                       open_auto := "Valves Data".R14_XV09.CMD,
                       open_man := "Valves Data".R14_XV09.MCMD,
                       fbk_open := "A/SSR_014_XV655_OFB",
                       fbk_close := "A/SSR_014_XV655_CFB",
                       reset := "Valves Data".R14_XV09.RESET OR "R14_DATA".R14.Reset,
                       intl := NOT "DI_INPUTS".R14_INPUTS_RUA.EMG_PB,
                       Mon_En := 1,
                       mon_sp := "Valves Data".R14_XV09.MON_TIME,
                       SEMI := "Valves Data".SEMI_AUTO.R14,
                       "open/close" => "A/SSR_014_XV655_CMD",
                       FAIL_TO_OPEN => "Valves Data".R14_VALVE_FAULT.XV09_FAIL_TO_OPEN,
                       FAIL_TO_CLOSE => "Valves Data".R14_VALVE_FAULT.XV09_FAIL_TO_CLOSE,
                       status => "Valves Data".R14_XV09.STATUS);
   END_IF;
END_REGION

REGION Network 152: R14_XV10
   RUNG wire#powerrail
      Contact( "AlwaysTRUE" )
      #valve_R14_XV10(reset := wire#w1, intl := wire#w2, "auto/manual" := "Valves Data"."A/M".R14, open_auto := "Valves Data".R14_XV10.CMD, open_man := "Valves Data".R14_XV10.MCMD, fbk_open := "A/SSR_014_XV401_OFB", fbk_close := "A/SSR_014_XV401_CFB", Mon_En := 1, mon_sp := "Valves Data".R14_XV10.MON_TIME, SEMI := "Valves Data".SEMI_AUTO.R14, SIM :=, "open/close" => "A/SSR_014_XV401_CMD", FAIL_TO_OPEN => "Valves Data".R14_VALVE_FAULT.XV010_FAIL_TO_OPEN, FAIL_TO_CLOSE => "Valves Data".R14_VALVE_FAULT.XV10_FAIL_TO_CLOSE, status => "Valves Data".R14_XV10.STATUS)
   END_RUNG
   RUNG wire#powerrail
      Contact( "Valves Data".R14_XV10.RESET )
   END_RUNG wire#w1
   RUNG wire#powerrail
      Contact( "R14_DATA".R14.Reset )
   END_RUNG wire#w1
   RUNG wire#powerrail
      I_Contact( "DI_INPUTS".R14_INPUTS_RUA.EMG_PB )
   END_RUNG wire#w2
   // the same network as SCL:
   IF "AlwaysTRUE" THEN
       #valve_R14_XV10("auto/manual" := "Valves Data"."A/M".R14,   // "valve"
                       open_auto := "Valves Data".R14_XV10.CMD,
                       open_man := "Valves Data".R14_XV10.MCMD,
                       fbk_open := "A/SSR_014_XV401_OFB",
                       fbk_close := "A/SSR_014_XV401_CFB",
                       reset := "Valves Data".R14_XV10.RESET OR "R14_DATA".R14.Reset,
                       intl := NOT "DI_INPUTS".R14_INPUTS_RUA.EMG_PB,
                       Mon_En := 1,
                       mon_sp := "Valves Data".R14_XV10.MON_TIME,
                       SEMI := "Valves Data".SEMI_AUTO.R14,
                       "open/close" => "A/SSR_014_XV401_CMD",
                       FAIL_TO_OPEN => "Valves Data".R14_VALVE_FAULT.XV010_FAIL_TO_OPEN,
                       FAIL_TO_CLOSE => "Valves Data".R14_VALVE_FAULT.XV10_FAIL_TO_CLOSE,
                       status => "Valves Data".R14_XV10.STATUS);
   END_IF;
END_REGION

REGION Network 153: ****REACTOR_15****
END_REGION

REGION Network 154: R15_XV01
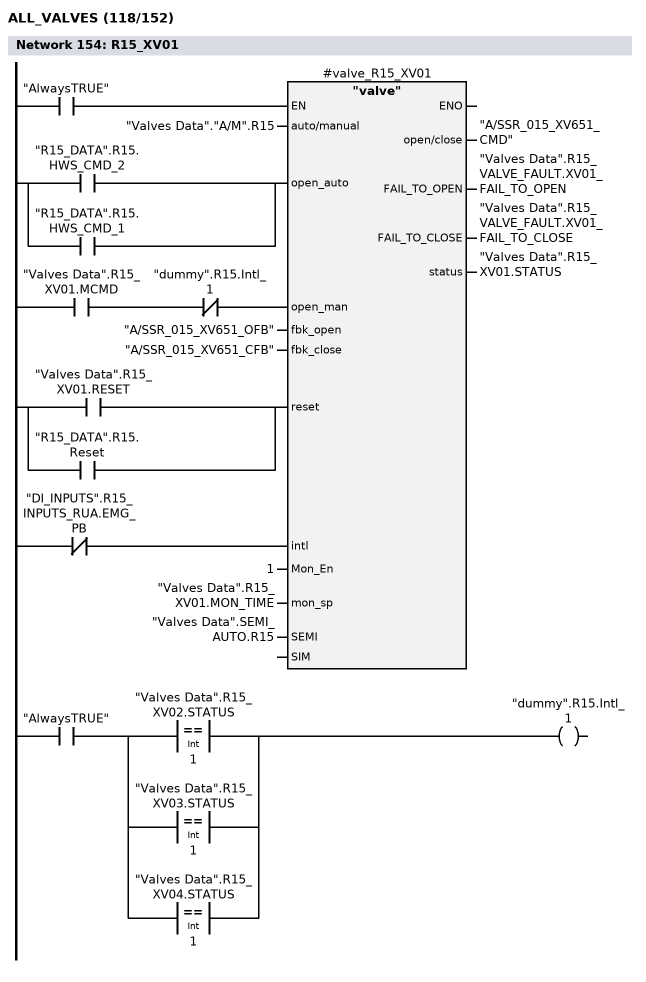
   RUNG wire#powerrail
      Contact( "AlwaysTRUE" )
      #valve_R15_XV01(open_auto := wire#w1, open_man := wire#w2, reset := wire#w3, intl := wire#w4, "auto/manual" := "Valves Data"."A/M".R15, fbk_open := "A/SSR_015_XV651_OFB", fbk_close := "A/SSR_015_XV651_CFB", Mon_En := 1, mon_sp := "Valves Data".R15_XV01.MON_TIME, SEMI := "Valves Data".SEMI_AUTO.R15, SIM :=, "open/close" => "A/SSR_015_XV651_CMD", FAIL_TO_OPEN => "Valves Data".R15_VALVE_FAULT.XV01_FAIL_TO_OPEN, FAIL_TO_CLOSE => "Valves Data".R15_VALVE_FAULT.XV01_FAIL_TO_CLOSE, status => "Valves Data".R15_XV01.STATUS)
   END_RUNG
   RUNG wire#powerrail
      Contact( "R15_DATA".R15.HWS_CMD_2 )
   END_RUNG wire#w1
   RUNG wire#powerrail
      Contact( "R15_DATA".R15.HWS_CMD_1 )
   END_RUNG wire#w1
   RUNG wire#powerrail
      Contact( "Valves Data".R15_XV01.MCMD )
      I_Contact( "dummy".R15.Intl_1 )
   END_RUNG wire#w2
   RUNG wire#powerrail
      Contact( "Valves Data".R15_XV01.RESET )
   END_RUNG wire#w3
   RUNG wire#powerrail
      Contact( "R15_DATA".R15.Reset )
   END_RUNG wire#w3
   RUNG wire#powerrail
      I_Contact( "DI_INPUTS".R15_INPUTS_RUA.EMG_PB )
   END_RUNG wire#w4
   RUNG wire#powerrail
      Contact( "AlwaysTRUE" )
      wire#w5
      { S7_Templates := "SrcType := Int" } EQ_Contact(in1 := "Valves Data".R15_XV02.STATUS, in2 := 1)
      wire#w6
      Coil( "dummy".R15.Intl_1 )
   END_RUNG
   RUNG wire#w5
      { S7_Templates := "SrcType := Int" } EQ_Contact(in1 := "Valves Data".R15_XV03.STATUS, in2 := 1)
   END_RUNG wire#w6
   RUNG wire#w5
      { S7_Templates := "SrcType := Int" } EQ_Contact(in1 := "Valves Data".R15_XV04.STATUS, in2 := 1)
   END_RUNG wire#w6
   // the same network as SCL:
   IF "AlwaysTRUE" THEN
       #valve_R15_XV01("auto/manual" := "Valves Data"."A/M".R15,   // "valve"
                       open_auto := "R15_DATA".R15.HWS_CMD_2 OR "R15_DATA".R15.HWS_CMD_1,
                       open_man := "Valves Data".R15_XV01.MCMD AND NOT "dummy".R15.Intl_1,
                       fbk_open := "A/SSR_015_XV651_OFB",
                       fbk_close := "A/SSR_015_XV651_CFB",
                       reset := "Valves Data".R15_XV01.RESET OR "R15_DATA".R15.Reset,
                       intl := NOT "DI_INPUTS".R15_INPUTS_RUA.EMG_PB,
                       Mon_En := 1,
                       mon_sp := "Valves Data".R15_XV01.MON_TIME,
                       SEMI := "Valves Data".SEMI_AUTO.R15,
                       "open/close" => "A/SSR_015_XV651_CMD",
                       FAIL_TO_OPEN => "Valves Data".R15_VALVE_FAULT.XV01_FAIL_TO_OPEN,
                       FAIL_TO_CLOSE => "Valves Data".R15_VALVE_FAULT.XV01_FAIL_TO_CLOSE,
                       status => "Valves Data".R15_XV01.STATUS);
   END_IF;
   "dummy".R15.Intl_1 := "AlwaysTRUE" AND (("Valves Data".R15_XV02.STATUS = 1) OR ("Valves Data".R15_XV03.STATUS = 1) OR ("Valves Data".R15_XV04.STATUS = 1));
END_REGION

REGION Network 155: R15_XV02
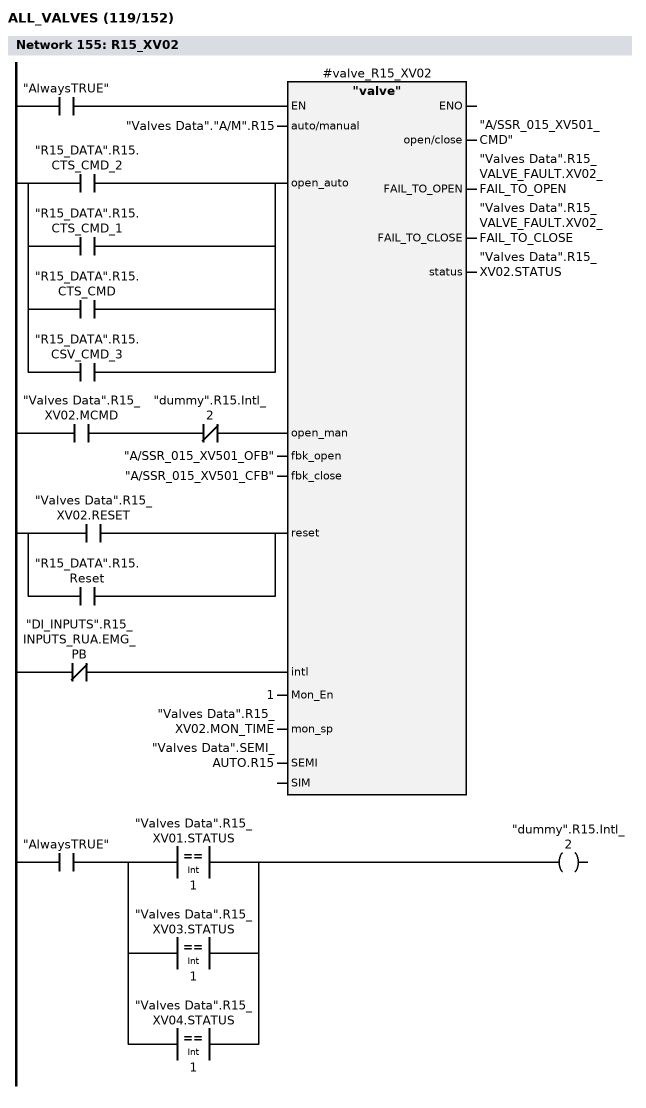
   RUNG wire#powerrail
      Contact( "AlwaysTRUE" )
      #valve_R15_XV02(open_auto := wire#w1, open_man := wire#w2, reset := wire#w3, intl := wire#w4, "auto/manual" := "Valves Data"."A/M".R15, fbk_open := "A/SSR_015_XV501_OFB", fbk_close := "A/SSR_015_XV501_CFB", Mon_En := 1, mon_sp := "Valves Data".R15_XV02.MON_TIME, SEMI := "Valves Data".SEMI_AUTO.R15, SIM :=, "open/close" => "A/SSR_015_XV501_CMD", FAIL_TO_OPEN => "Valves Data".R15_VALVE_FAULT.XV02_FAIL_TO_OPEN, FAIL_TO_CLOSE => "Valves Data".R15_VALVE_FAULT.XV02_FAIL_TO_CLOSE, status => "Valves Data".R15_XV02.STATUS)
   END_RUNG
   RUNG wire#powerrail
      Contact( "R15_DATA".R15.CTS_CMD_2 )
   END_RUNG wire#w1
   RUNG wire#powerrail
      Contact( "R15_DATA".R15.CTS_CMD_1 )
   END_RUNG wire#w1
   RUNG wire#powerrail
      Contact( "R15_DATA".R15.CTS_CMD )
   END_RUNG wire#w1
   RUNG wire#powerrail
      Contact( "R15_DATA".R15.CSV_CMD_3 )
   END_RUNG wire#w1
   RUNG wire#powerrail
      Contact( "Valves Data".R15_XV02.MCMD )
      I_Contact( "dummy".R15.Intl_2 )
   END_RUNG wire#w2
   RUNG wire#powerrail
      Contact( "Valves Data".R15_XV02.RESET )
   END_RUNG wire#w3
   RUNG wire#powerrail
      Contact( "R15_DATA".R15.Reset )
   END_RUNG wire#w3
   RUNG wire#powerrail
      I_Contact( "DI_INPUTS".R15_INPUTS_RUA.EMG_PB )
   END_RUNG wire#w4
   RUNG wire#powerrail
      Contact( "AlwaysTRUE" )
      wire#w5
      { S7_Templates := "SrcType := Int" } EQ_Contact(in1 := "Valves Data".R15_XV01.STATUS, in2 := 1)
      wire#w6
      Coil( "dummy".R15.Intl_2 )
   END_RUNG
   RUNG wire#w5
      { S7_Templates := "SrcType := Int" } EQ_Contact(in1 := "Valves Data".R15_XV03.STATUS, in2 := 1)
   END_RUNG wire#w6
   RUNG wire#w5
      { S7_Templates := "SrcType := Int" } EQ_Contact(in1 := "Valves Data".R15_XV04.STATUS, in2 := 1)
   END_RUNG wire#w6
   // the same network as SCL:
   IF "AlwaysTRUE" THEN
       #valve_R15_XV02("auto/manual" := "Valves Data"."A/M".R15,   // "valve"
                       open_auto := "R15_DATA".R15.CTS_CMD_2 OR "R15_DATA".R15.CTS_CMD_1 OR "R15_DATA".R15.CTS_CMD OR "R15_DATA".R15.CSV_CMD_3,
                       open_man := "Valves Data".R15_XV02.MCMD AND NOT "dummy".R15.Intl_2,
                       fbk_open := "A/SSR_015_XV501_OFB",
                       fbk_close := "A/SSR_015_XV501_CFB",
                       reset := "Valves Data".R15_XV02.RESET OR "R15_DATA".R15.Reset,
                       intl := NOT "DI_INPUTS".R15_INPUTS_RUA.EMG_PB,
                       Mon_En := 1,
                       mon_sp := "Valves Data".R15_XV02.MON_TIME,
                       SEMI := "Valves Data".SEMI_AUTO.R15,
                       "open/close" => "A/SSR_015_XV501_CMD",
                       FAIL_TO_OPEN => "Valves Data".R15_VALVE_FAULT.XV02_FAIL_TO_OPEN,
                       FAIL_TO_CLOSE => "Valves Data".R15_VALVE_FAULT.XV02_FAIL_TO_CLOSE,
                       status => "Valves Data".R15_XV02.STATUS);
   END_IF;
   "dummy".R15.Intl_2 := "AlwaysTRUE" AND (("Valves Data".R15_XV01.STATUS = 1) OR ("Valves Data".R15_XV03.STATUS = 1) OR ("Valves Data".R15_XV04.STATUS = 1));
END_REGION

REGION Network 156: R15_XV03
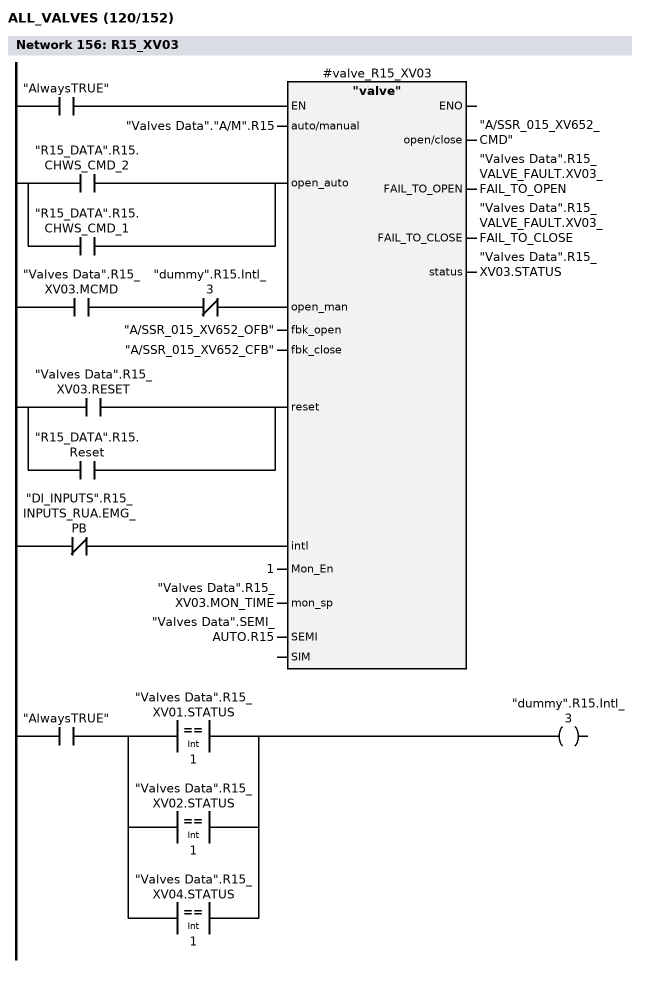
   RUNG wire#powerrail
      Contact( "AlwaysTRUE" )
      #valve_R15_XV03(open_auto := wire#w1, open_man := wire#w2, reset := wire#w3, intl := wire#w4, "auto/manual" := "Valves Data"."A/M".R15, fbk_open := "A/SSR_015_XV652_OFB", fbk_close := "A/SSR_015_XV652_CFB", Mon_En := 1, mon_sp := "Valves Data".R15_XV03.MON_TIME, SEMI := "Valves Data".SEMI_AUTO.R15, SIM :=, "open/close" => "A/SSR_015_XV652_CMD", FAIL_TO_OPEN => "Valves Data".R15_VALVE_FAULT.XV03_FAIL_TO_OPEN, FAIL_TO_CLOSE => "Valves Data".R15_VALVE_FAULT.XV03_FAIL_TO_CLOSE, status => "Valves Data".R15_XV03.STATUS)
   END_RUNG
   RUNG wire#powerrail
      Contact( "R15_DATA".R15.CHWS_CMD_2 )
   END_RUNG wire#w1
   RUNG wire#powerrail
      Contact( "R15_DATA".R15.CHWS_CMD_1 )
   END_RUNG wire#w1
   RUNG wire#powerrail
      Contact( "Valves Data".R15_XV03.MCMD )
      I_Contact( "dummy".R15.Intl_3 )
   END_RUNG wire#w2
   RUNG wire#powerrail
      Contact( "Valves Data".R15_XV03.RESET )
   END_RUNG wire#w3
   RUNG wire#powerrail
      Contact( "R15_DATA".R15.Reset )
   END_RUNG wire#w3
   RUNG wire#powerrail
      I_Contact( "DI_INPUTS".R15_INPUTS_RUA.EMG_PB )
   END_RUNG wire#w4
   RUNG wire#powerrail
      Contact( "AlwaysTRUE" )
      wire#w5
      { S7_Templates := "SrcType := Int" } EQ_Contact(in1 := "Valves Data".R15_XV01.STATUS, in2 := 1)
      wire#w6
      Coil( "dummy".R15.Intl_3 )
   END_RUNG
   RUNG wire#w5
      { S7_Templates := "SrcType := Int" } EQ_Contact(in1 := "Valves Data".R15_XV02.STATUS, in2 := 1)
   END_RUNG wire#w6
   RUNG wire#w5
      { S7_Templates := "SrcType := Int" } EQ_Contact(in1 := "Valves Data".R15_XV04.STATUS, in2 := 1)
   END_RUNG wire#w6
   // the same network as SCL:
   IF "AlwaysTRUE" THEN
       #valve_R15_XV03("auto/manual" := "Valves Data"."A/M".R15,   // "valve"
                       open_auto := "R15_DATA".R15.CHWS_CMD_2 OR "R15_DATA".R15.CHWS_CMD_1,
                       open_man := "Valves Data".R15_XV03.MCMD AND NOT "dummy".R15.Intl_3,
                       fbk_open := "A/SSR_015_XV652_OFB",
                       fbk_close := "A/SSR_015_XV652_CFB",
                       reset := "Valves Data".R15_XV03.RESET OR "R15_DATA".R15.Reset,
                       intl := NOT "DI_INPUTS".R15_INPUTS_RUA.EMG_PB,
                       Mon_En := 1,
                       mon_sp := "Valves Data".R15_XV03.MON_TIME,
                       SEMI := "Valves Data".SEMI_AUTO.R15,
                       "open/close" => "A/SSR_015_XV652_CMD",
                       FAIL_TO_OPEN => "Valves Data".R15_VALVE_FAULT.XV03_FAIL_TO_OPEN,
                       FAIL_TO_CLOSE => "Valves Data".R15_VALVE_FAULT.XV03_FAIL_TO_CLOSE,
                       status => "Valves Data".R15_XV03.STATUS);
   END_IF;
   "dummy".R15.Intl_3 := "AlwaysTRUE" AND (("Valves Data".R15_XV01.STATUS = 1) OR ("Valves Data".R15_XV02.STATUS = 1) OR ("Valves Data".R15_XV04.STATUS = 1));
END_REGION

REGION Network 157: R15_XV04
